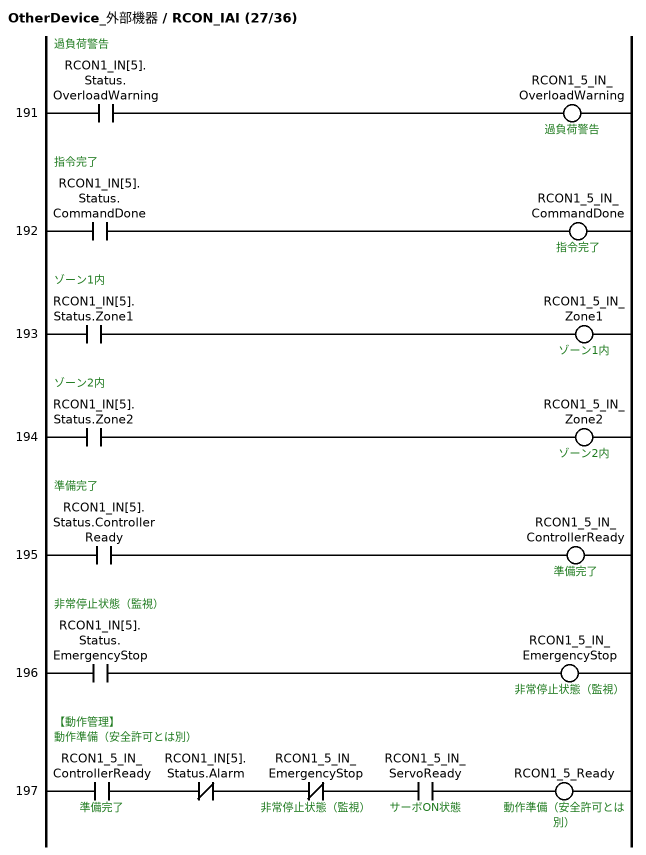
(* [picture p72: OtherDevice_外部機器 / RCON_IAI, rungs 191-197] *)
(* Rung 191: 過負荷警告 *)
RCON1_5_IN_OverloadWarning := RCON1_IN[5].Status.OverloadWarning;
(* Rung 192: 指令完了 *)
RCON1_5_IN_CommandDone := RCON1_IN[5].Status.CommandDone;
(* Rung 193: ゾーン1内 *)
RCON1_5_IN_Zone1 := RCON1_IN[5].Status.Zone1;
(* Rung 194: ゾーン2内 *)
RCON1_5_IN_Zone2 := RCON1_IN[5].Status.Zone2;
(* Rung 195: 準備完了 *)
RCON1_5_IN_ControllerReady := RCON1_IN[5].Status.ControllerReady;
(* Rung 196: 非常停止状態（監視） *)
RCON1_5_IN_EmergencyStop := RCON1_IN[5].Status.EmergencyStop;
(* Rung 197: 【動作管理】 / 動作準備（安全許可とは別） *)
RCON1_5_Ready := RCON1_5_IN_ControllerReady AND NOT RCON1_IN[5].Status.Alarm AND NOT RCON1_5_IN_EmergencyStop AND RCON1_5_IN_ServoReady;

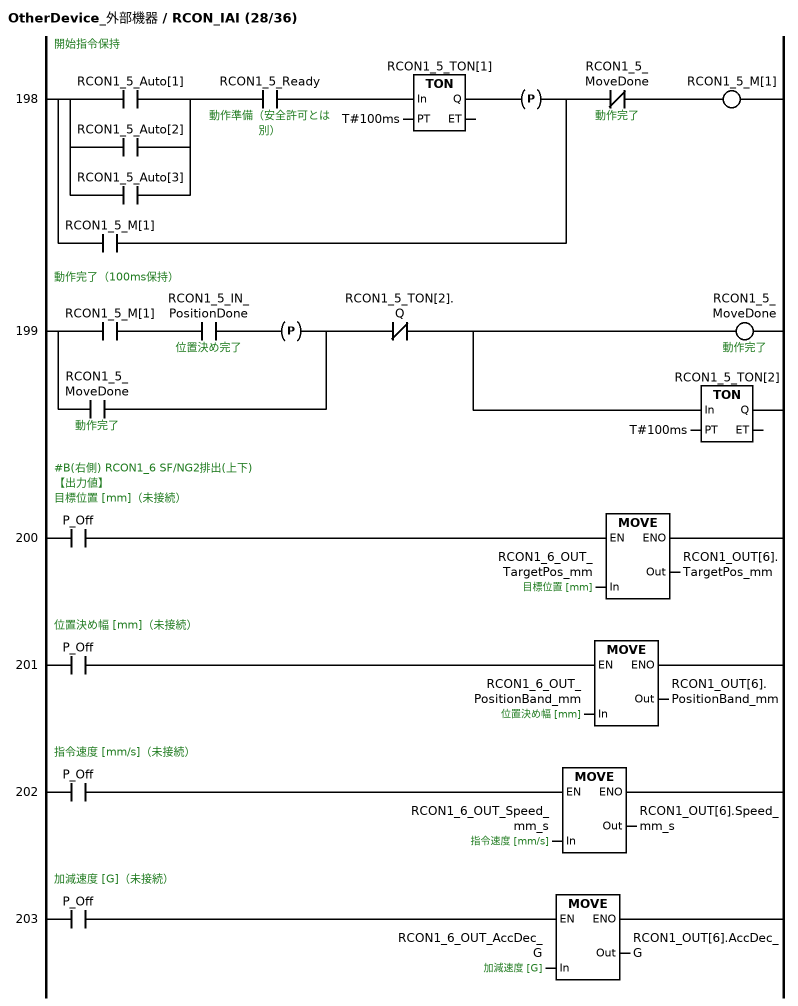
(* Rung 198: 開始指令保持 *)
RCON1_5_TON[1](In := (RCON1_5_Auto[1] OR RCON1_5_Auto[2] OR RCON1_5_Auto[3]) AND RCON1_5_Ready, PT := T#100ms);
_e18(CLK := RCON1_5_TON[1].Q);
RCON1_5_M[1] := (_e18.Q OR RCON1_5_M[1]) AND NOT RCON1_5_MoveDone;
(* Rung 199: 動作完了（100ms保持） *)
_e19(CLK := RCON1_5_M[1] AND RCON1_5_IN_PositionDone);
_p20 := (_e19.Q OR RCON1_5_MoveDone) AND NOT RCON1_5_TON[2].Q;
RCON1_5_MoveDone := _p20;
RCON1_5_TON[2](In := _p20, PT := T#100ms);
(* Rung 200: #B(右側) RCON1_6 SF/NG2排出(上下) / 【出力値】 / 目標位置 [mm]（未接続） *)
IF P_Off THEN RCON1_OUT[6].TargetPos_mm := RCON1_6_OUT_TargetPos_mm; END_IF;
(* Rung 201: 位置決め幅 [mm]（未接続） *)
IF P_Off THEN RCON1_OUT[6].PositionBand_mm := RCON1_6_OUT_PositionBand_mm; END_IF;
(* Rung 202: 指令速度 [mm/s]（未接続） *)
IF P_Off THEN RCON1_OUT[6].Speed_mm_s := RCON1_6_OUT_Speed_mm_s; END_IF;
(* Rung 203: 加減速度 [G]（未接続） *)
IF P_Off THEN RCON1_OUT[6].AccDec_G := RCON1_6_OUT_AccDec_G; END_IF;

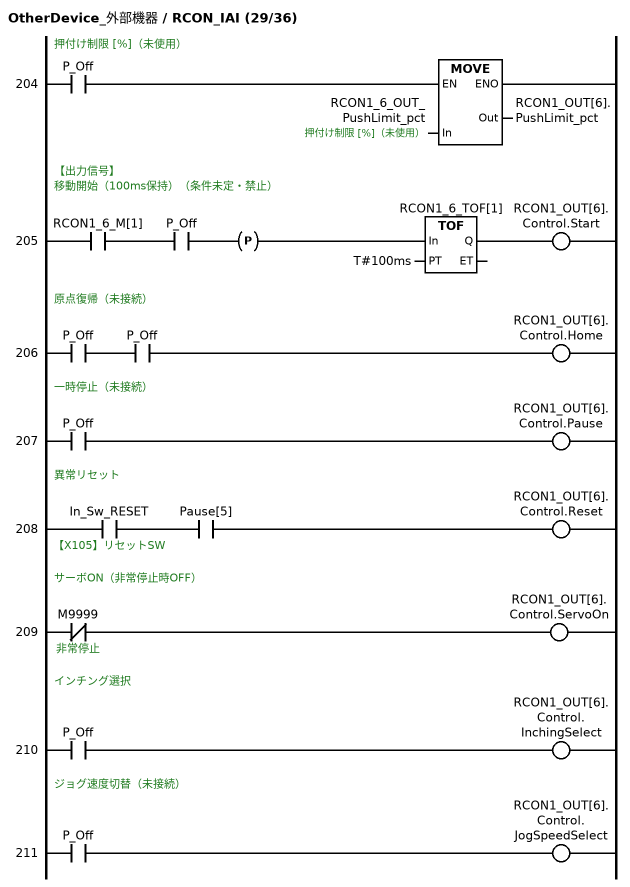
(* Rung 204: 押付け制限 [%]（未使用） *)
IF P_Off THEN RCON1_OUT[6].PushLimit_pct := RCON1_6_OUT_PushLimit_pct; END_IF;
(* Rung 205: 【出力信号】 / 移動開始（100ms保持）（条件未定・禁止） *)
_e21(CLK := RCON1_6_M[1] AND P_Off);
RCON1_6_TOF[1](In := _e21.Q, PT := T#100ms);
RCON1_OUT[6].Control.Start := RCON1_6_TOF[1].Q;
(* Rung 206: 原点復帰（未接続） *)
RCON1_OUT[6].Control.Home := P_Off AND P_Off;
(* Rung 207: 一時停止（未接続） *)
RCON1_OUT[6].Control.Pause := P_Off;
(* Rung 208: 異常リセット *)
RCON1_OUT[6].Control.Reset := In_Sw_RESET AND Pause[5];
(* Rung 209: サーボON（非常停止時OFF） *)
RCON1_OUT[6].Control.ServoOn := NOT M9999;
(* Rung 210: インチング選択 *)
RCON1_OUT[6].Control.InchingSelect := P_Off;
(* Rung 211: ジョグ速度切替（未接続） *)
RCON1_OUT[6].Control.JogSpeedSelect := P_Off;

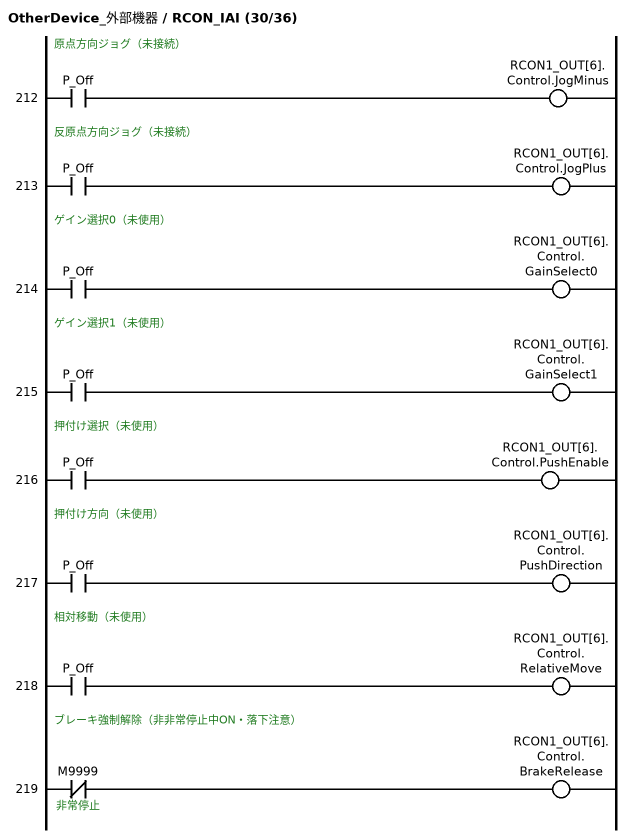
(* Rung 212: 原点方向ジョグ（未接続） *)
RCON1_OUT[6].Control.JogMinus := P_Off;
(* Rung 213: 反原点方向ジョグ（未接続） *)
RCON1_OUT[6].Control.JogPlus := P_Off;
(* Rung 214: ゲイン選択0（未使用） *)
RCON1_OUT[6].Control.GainSelect0 := P_Off;
(* Rung 215: ゲイン選択1（未使用） *)
RCON1_OUT[6].Control.GainSelect1 := P_Off;
(* Rung 216: 押付け選択（未使用） *)
RCON1_OUT[6].Control.PushEnable := P_Off;
(* Rung 217: 押付け方向（未使用） *)
RCON1_OUT[6].Control.PushDirection := P_Off;
(* Rung 218: 相対移動（未使用） *)
RCON1_OUT[6].Control.RelativeMove := P_Off;
(* Rung 219: ブレーキ強制解除（非非常停止中ON・落下注意） *)
RCON1_OUT[6].Control.BrakeRelease := NOT M9999;

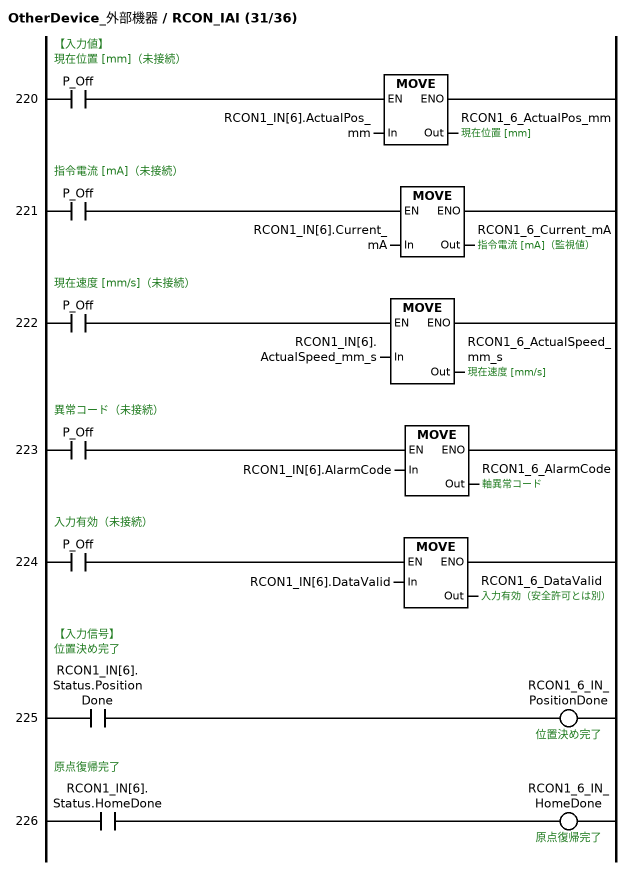
(* Rung 220: 【入力値】 / 現在位置 [mm]（未接続） *)
IF P_Off THEN RCON1_6_ActualPos_mm := RCON1_IN[6].ActualPos_mm; END_IF;
(* Rung 221: 指令電流 [mA]（未接続） *)
IF P_Off THEN RCON1_6_Current_mA := RCON1_IN[6].Current_mA; END_IF;
(* Rung 222: 現在速度 [mm/s]（未接続） *)
IF P_Off THEN RCON1_6_ActualSpeed_mm_s := RCON1_IN[6].ActualSpeed_mm_s; END_IF;
(* Rung 223: 異常コード（未接続） *)
IF P_Off THEN RCON1_6_AlarmCode := RCON1_IN[6].AlarmCode; END_IF;
(* Rung 224: 入力有効（未接続） *)
IF P_Off THEN RCON1_6_DataValid := RCON1_IN[6].DataValid; END_IF;
(* Rung 225: 【入力信号】 / 位置決め完了 *)
RCON1_6_IN_PositionDone := RCON1_IN[6].Status.PositionDone;
(* Rung 226: 原点復帰完了 *)
RCON1_6_IN_HomeDone := RCON1_IN[6].Status.HomeDone;

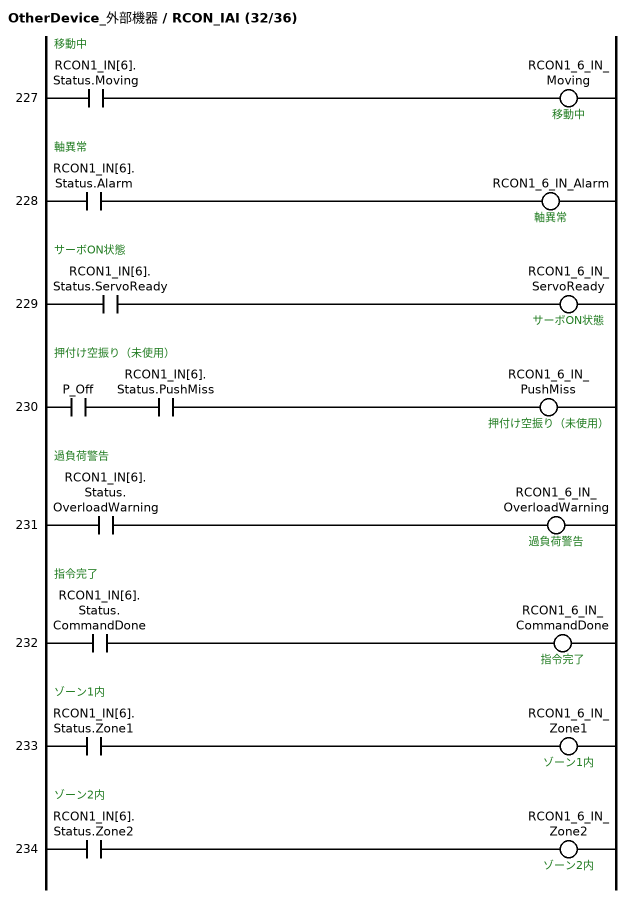
(* Rung 227: 移動中 *)
RCON1_6_IN_Moving := RCON1_IN[6].Status.Moving;
(* Rung 228: 軸異常 *)
RCON1_6_IN_Alarm := RCON1_IN[6].Status.Alarm;
(* Rung 229: サーボON状態 *)
RCON1_6_IN_ServoReady := RCON1_IN[6].Status.ServoReady;
(* Rung 230: 押付け空振り（未使用） *)
RCON1_6_IN_PushMiss := P_Off AND RCON1_IN[6].Status.PushMiss;
(* Rung 231: 過負荷警告 *)
RCON1_6_IN_OverloadWarning := RCON1_IN[6].Status.OverloadWarning;
(* Rung 232: 指令完了 *)
RCON1_6_IN_CommandDone := RCON1_IN[6].Status.CommandDone;
(* Rung 233: ゾーン1内 *)
RCON1_6_IN_Zone1 := RCON1_IN[6].Status.Zone1;
(* Rung 234: ゾーン2内 *)
RCON1_6_IN_Zone2 := RCON1_IN[6].Status.Zone2;

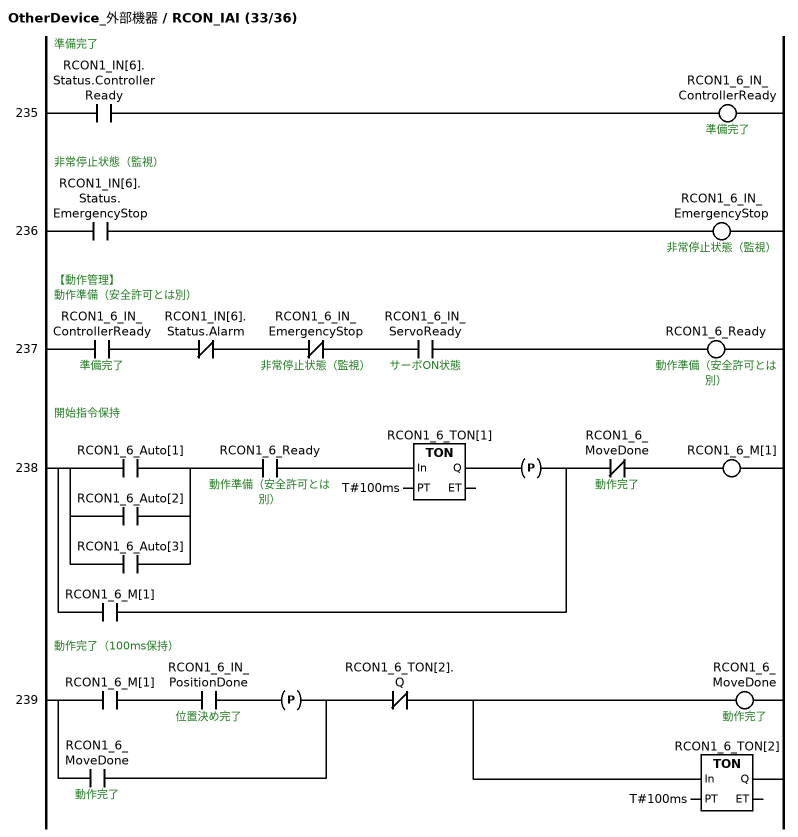
(* Rung 235: 準備完了 *)
RCON1_6_IN_ControllerReady := RCON1_IN[6].Status.ControllerReady;
(* Rung 236: 非常停止状態（監視） *)
RCON1_6_IN_EmergencyStop := RCON1_IN[6].Status.EmergencyStop;
(* Rung 237: 【動作管理】 / 動作準備（安全許可とは別） *)
RCON1_6_Ready := RCON1_6_IN_ControllerReady AND NOT RCON1_IN[6].Status.Alarm AND NOT RCON1_6_IN_EmergencyStop AND RCON1_6_IN_ServoReady;
(* Rung 238: 開始指令保持 *)
RCON1_6_TON[1](In := (RCON1_6_Auto[1] OR RCON1_6_Auto[2] OR RCON1_6_Auto[3]) AND RCON1_6_Ready, PT := T#100ms);
_e22(CLK := RCON1_6_TON[1].Q);
RCON1_6_M[1] := (_e22.Q OR RCON1_6_M[1]) AND NOT RCON1_6_MoveDone;
(* Rung 239: 動作完了（100ms保持） *)
_e23(CLK := RCON1_6_M[1] AND RCON1_6_IN_PositionDone);
_p24 := (_e23.Q OR RCON1_6_MoveDone) AND NOT RCON1_6_TON[2].Q;
RCON1_6_MoveDone := _p24;
RCON1_6_TON[2](In := _p24, PT := T#100ms);

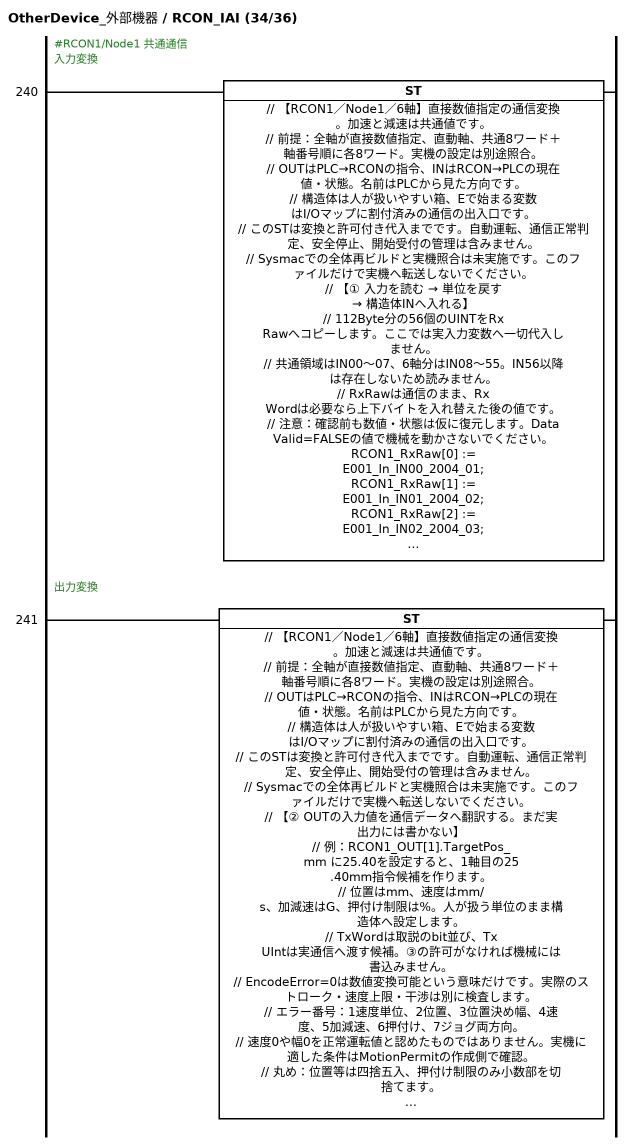
(* Rung 240: #RCON1/Node1 共通通信 / 入力変換 *)
// 【RCON1／Node1／6軸】直接数値指定の通信変換。加速と減速は共通値です。
// 前提：全軸が直接数値指定、直動軸、共通8ワード＋軸番号順に各8ワード。実機の設定は別途照合。
// OUTはPLC→RCONの指令、INはRCON→PLCの現在値・状態。名前はPLCから見た方向です。
// 構造体は人が扱いやすい箱、Eで始まる変数はI/Oマップに割付済みの通信の出入口です。
// このSTは変換と許可付き代入までです。自動運転、通信正常判定、安全停止、開始受付の管理は含みません。
// Sysmacでの全体再ビルドと実機照合は未実施です。このファイルだけで実機へ転送しないでください。
// 【① 入力を読む → 単位を戻す → 構造体INへ入れる】
// 112Byte分の56個のUINTをRxRawへコピーします。ここでは実入力変数へ一切代入しません。
// 共通領域はIN00～07、6軸分はIN08～55。IN56以降は存在しないため読みません。
// RxRawは通信のまま、RxWordは必要なら上下バイトを入れ替えた後の値です。
// 注意：確認前も数値・状態は仮に復元します。DataValid=FALSEの値で機械を動かさないでください。
RCON1_RxRaw[0] := E001_In_IN00_2004_01;
RCON1_RxRaw[1] := E001_In_IN01_2004_02;
RCON1_RxRaw[2] := E001_In_IN02_2004_03;
RCON1_RxRaw[3] := E001_In_IN03_2004_04;
RCON1_RxRaw[4] := E001_In_IN04_2004_05;
RCON1_RxRaw[5] := E001_In_IN05_2004_06;
RCON1_RxRaw[6] := E001_In_IN06_2004_07;
RCON1_RxRaw[7] := E001_In_IN07_2004_08;
RCON1_RxRaw[8] := E001_In_IN08_2004_09;
RCON1_RxRaw[9] := E001_In_IN09_2004_0A;
RCON1_RxRaw[10] := E001_In_IN10_2004_0B;
RCON1_RxRaw[11] := E001_In_IN11_2004_0C;
RCON1_RxRaw[12] := E001_In_IN12_2004_0D;
RCON1_RxRaw[13] := E001_In_IN13_2004_0E;
RCON1_RxRaw[14] := E001_In_IN14_2004_0F;
RCON1_RxRaw[15] := E001_In_IN15_2004_10;
RCON1_RxRaw[16] := E001_In_IN16_2004_11;
RCON1_RxRaw[17] := E001_In_IN17_2004_12;
RCON1_RxRaw[18] := E001_In_IN18_2004_13;
RCON1_RxRaw[19] := E001_In_IN19_2004_14;
RCON1_RxRaw[20] := E001_In_IN20_2004_15;
RCON1_RxRaw[21] := E001_In_IN21_2004_16;
RCON1_RxRaw[22] := E001_In_IN22_2004_17;
RCON1_RxRaw[23] := E001_In_IN23_2004_18;
RCON1_RxRaw[24] := E001_In_IN24_2004_19;
RCON1_RxRaw[25] := E001_In_IN25_2004_1A;
RCON1_RxRaw[26] := E001_In_IN26_2004_1B;
RCON1_RxRaw[27] := E001_In_IN27_2004_1C;
RCON1_RxRaw[28] := E001_In_IN28_2004_1D;
RCON1_RxRaw[29] := E001_In_IN29_2004_1E;
RCON1_RxRaw[30] := E001_In_IN30_2004_1F;
RCON1_RxRaw[31] := E001_In_IN31_2004_20;
RCON1_RxRaw[32] := E001_In_IN32_2004_21;
RCON1_RxRaw[33] := E001_In_IN33_2004_22;
RCON1_RxRaw[34] := E001_In_IN34_2004_23;
RCON1_RxRaw[35] := E001_In_IN35_2004_24;
RCON1_RxRaw[36] := E001_In_IN36_2004_25;
RCON1_RxRaw[37] := E001_In_IN37_2004_26;
RCON1_RxRaw[38] := E001_In_IN38_2004_27;
RCON1_RxRaw[39] := E001_In_IN39_2004_28;
RCON1_RxRaw[40] := E001_In_IN40_2004_29;
RCON1_RxRaw[41] := E001_In_IN41_2004_2A;
RCON1_RxRaw[42] := E001_In_IN42_2004_2B;
RCON1_RxRaw[43] := E001_In_IN43_2004_2C;
RCON1_RxRaw[44] := E001_In_IN44_2004_2D;
RCON1_RxRaw[45] := E001_In_IN45_2004_2E;
RCON1_RxRaw[46] := E001_In_IN46_2004_2F;
RCON1_RxRaw[47] := E001_In_IN47_2004_30;
RCON1_RxRaw[48] := E001_In_IN48_2004_31;
RCON1_RxRaw[49] := E001_In_IN49_2004_32;
RCON1_RxRaw[50] := E001_In_IN50_2004_33;
RCON1_RxRaw[51] := E001_In_IN51_2004_34;
RCON1_RxRaw[52] := E001_In_IN52_2004_35;
RCON1_RxRaw[53] := E001_In_IN53_2004_36;
RCON1_RxRaw[54] := E001_In_IN54_2004_37;
RCON1_RxRaw[55] := E001_In_IN55_2004_38;
// 取説の論理ワードへ正規化。Swapは1ワード内の上下バイト交換です。
// SwapBytesは推測で設定せず、既知の位置とbitで実機照合してください。
FOR ConvWordIndex := INT#0 TO INT#55 DO
    RCON1_RxWord[ConvWordIndex] := UINT_TO_WORD(RCON1_RxRaw[ConvWordIndex]);
    IF RCON1_SwapBytes THEN
        RCON1_RxWord[ConvWordIndex] := Swap(RCON1_RxWord[ConvWordIndex]);
    END_IF;
END_FOR;

ConvUnitOK := (RCON1_SpeedUnit_mm_s = LREAL#1.0) OR
              (RCON1_SpeedUnit_mm_s = LREAL#0.1);

// 【①-2 共通状態】IN00はユニット全体、IN01は各軸のリンク情報です。
// TestABit(ワード, bit番号)は、そのスイッチがONかをBOOLで取り出す命令です。
// 例：IN01のb0は軸No.0→配列[1]、b1は軸No.1→配列[2]。配列番号と実機軸番号は1違います。
// 共通固定領域。ここで使うbit番号は取説の論理bitです（MJ0384 6-24～6-25）。
RCON1_GwRun := TestABit(RCON1_RxWord[0], USINT#15);
RCON1_GwControllerCommLatch := TestABit(RCON1_RxWord[0], USINT#14);
RCON1_GwAxisCommError := TestABit(RCON1_RxWord[0], USINT#13);
RCON1_GwManual := TestABit(RCON1_RxWord[0], USINT#12);
RCON1_GwHeavyAlarm := TestABit(RCON1_RxWord[0], USINT#11);
RCON1_GwLightAlarm := TestABit(RCON1_RxWord[0], USINT#10);
RCON1_GwSystemStop := TestABit(RCON1_RxWord[0], USINT#8);
RCON1_GwAlarmCode := WORD_TO_UINT(RCON1_RxWord[0] AND WORD#16#00FF);
FOR ConvWordIndex := INT#0 TO INT#4 DO
    RCON1_PowerStateRaw[ConvWordIndex] := RCON1_RxWord[ConvWordIndex + INT#2];
END_FOR;

// 【①-3 軸ごとに同じ読取りを繰り返す】
// FORは1～6軸を順番に処理します。ConvBaseはその軸の先頭番号です。
// 計算：8+(軸番号-1)×8。1軸目=8、2軸目=16、3軸目=24。先頭8ワードは共通領域です。
FOR ConvAxisIndex := INT#1 TO INT#6 DO
    ConvBase := INT#8 + (ConvAxisIndex - INT#1) * INT#8;
    RCON1_AxisLinked[ConvAxisIndex] :=
        TestABit(RCON1_RxWord[1], INT_TO_USINT(ConvAxisIndex - INT#1));

// 例：下位2540／上位0なら32bit値2540→25.40mm。
// 上位を16bit左に動かして下位とORで重ねます。SHLが左シフト、ORがビットの合成です。
// 負位置はDWORD_TO_DINTで符号を復元。下位62996／上位65535なら-2540→-25.40mm。
    // 現在位置：下位・上位を結合、符号付き32bitとして解釈、0.01mmをmmへ。
    ConvDWord := SHL(WORD_TO_DWORD(RCON1_RxWord[ConvBase + INT#1]), ULINT#16)
                 OR WORD_TO_DWORD(RCON1_RxWord[ConvBase]);
    RCON1_IN[ConvAxisIndex].ActualPos_mm :=
        DINT_TO_LREAL(DWORD_TO_DINT(ConvDWord)) * LREAL#0.01;

    // 電流：32bitのmA。RCON-PCでは指令電流であり、実測トルクではありません。
    ConvDWord := SHL(WORD_TO_DWORD(RCON1_RxWord[ConvBase + INT#3]), ULINT#16)
                 OR WORD_TO_DWORD(RCON1_RxWord[ConvBase + INT#2]);
    RCON1_IN[ConvAxisIndex].Current_mA := DWORD_TO_DINT(ConvDWord);

    // 現在速度：16bitの負数をINTとして読む。UINTのまま速度にしません。
    IF ConvUnitOK THEN
        RCON1_IN[ConvAxisIndex].ActualSpeed_mm_s :=
            INT_TO_LREAL(WORD_TO_INT(RCON1_RxWord[ConvBase + INT#4])) * RCON1_SpeedUnit_mm_s;
    END_IF;
    // 単位不明のとき速度は前値を保持し、DataValidはFALSEにします。
    // 軸内の+5ワードは予約のため値を使用しません。
    RCON1_IN[ConvAxisIndex].AlarmCode := WORD_TO_UINT(RCON1_RxWord[ConvBase + INT#6]);

// 例：Status.ServoReady=TRUEは「サーボON状態を受信した」という意味。
// OUT側Control.ServoOn=TRUEは「サーボONを要求する」という意味で、指令と結果を区別します。
    // 状態ワード：12個のBOOLへ分解。予約b6,b9～11は使いません。
    RCON1_IN[ConvAxisIndex].Status.PositionDone := TestABit(RCON1_RxWord[ConvBase + INT#7], USINT#0);
    RCON1_IN[ConvAxisIndex].Status.HomeDone := TestABit(RCON1_RxWord[ConvBase + INT#7], USINT#1);
    RCON1_IN[ConvAxisIndex].Status.Moving := TestABit(RCON1_RxWord[ConvBase + INT#7], USINT#2);
    RCON1_IN[ConvAxisIndex].Status.Alarm := TestABit(RCON1_RxWord[ConvBase + INT#7], USINT#3);
    RCON1_IN[ConvAxisIndex].Status.ServoReady := TestABit(RCON1_RxWord[ConvBase + INT#7], USINT#4);
    RCON1_IN[ConvAxisIndex].Status.PushMiss := TestABit(RCON1_RxWord[ConvBase + INT#7], USINT#5);
    RCON1_IN[ConvAxisIndex].Status.OverloadWarning := TestABit(RCON1_RxWord[ConvBase + INT#7], USINT#7);
    RCON1_IN[ConvAxisIndex].Status.CommandDone := TestABit(RCON1_RxWord[ConvBase + INT#7], USINT#8);
    RCON1_IN[ConvAxisIndex].Status.Zone1 := TestABit(RCON1_RxWord[ConvBase + INT#7], USINT#12);
    RCON1_IN[ConvAxisIndex].Status.Zone2 := TestABit(RCON1_RxWord[ConvBase + INT#7], USINT#13);
    RCON1_IN[ConvAxisIndex].Status.ControllerReady := TestABit(RCON1_RxWord[ConvBase + INT#7], USINT#14);
    RCON1_IN[ConvAxisIndex].Status.EmergencyStop := TestABit(RCON1_RxWord[ConvBase + INT#7], USINT#15);

    // DataValidは直接受信bitではなく、今回の内部設計で決めた内部判定です。
    // CommOKはCPUの実通信状態から別途作成。単にTRUE固定にしないでください。
    // DataValidは運転許可や安全保証ではありません。各異常・原点等は別途確認。
    RCON1_IN[ConvAxisIndex].DataValid := RCON1_CommOK AND RCON1_LayoutConfirmed
        AND RCON1_ByteOrderConfirmed AND ConvUnitOK AND RCON1_GwRun
        AND RCON1_AxisLinked[ConvAxisIndex] AND NOT RCON1_GwAxisCommError;
END_FOR;
(* Rung 241: 出力変換 *)
// 【RCON1／Node1／6軸】直接数値指定の通信変換。加速と減速は共通値です。
// 前提：全軸が直接数値指定、直動軸、共通8ワード＋軸番号順に各8ワード。実機の設定は別途照合。
// OUTはPLC→RCONの指令、INはRCON→PLCの現在値・状態。名前はPLCから見た方向です。
// 構造体は人が扱いやすい箱、Eで始まる変数はI/Oマップに割付済みの通信の出入口です。
// このSTは変換と許可付き代入までです。自動運転、通信正常判定、安全停止、開始受付の管理は含みません。
// Sysmacでの全体再ビルドと実機照合は未実施です。このファイルだけで実機へ転送しないでください。
// 【② OUTの入力値を通信データへ翻訳する。まだ実出力には書かない】
// 例：RCON1_OUT[1].TargetPos_mm に25.40を設定すると、1軸目の25.40mm指令候補を作ります。
// 位置はmm、速度はmm/s、加減速はG、押付け制限は%。人が扱う単位のまま構造体へ設定します。
// TxWordは取説のbit並び、TxUIntは実通信へ渡す候補。③の許可がなければ機械には書込みません。
// EncodeError=0は数値変換可能という意味だけです。実際のストローク・速度上限・干渉は別に検査します。
// エラー番号：1速度単位、2位置、3位置決め幅、4速度、5加減速、6押付け、7ジョグ両方向。
// 速度0や幅0を正常運転値と認めたものではありません。実機に適した条件はMotionPermitの作成側で確認。
// 丸め：位置等は四捨五入、押付け制限のみ小数部を切捨てます。

ConvUnitOK := (RCON1_SpeedUnit_mm_s = LREAL#1.0) OR
              (RCON1_SpeedUnit_mm_s = LREAL#0.1);

// 共通制御：MONは論理b15、RTEは論理b13。他のbitは0。
// MONを落とす処理を安全停止として扱わないでください。
RCON1_TxWord[0] := WORD#16#0000;
IF RCON1_GwMON_Request THEN
    RCON1_TxWord[0] := RCON1_TxWord[0] OR WORD#16#8000;
END_IF;
IF RCON1_GwRTE_Request THEN
    RCON1_TxWord[0] := RCON1_TxWord[0] OR WORD#16#2000;
END_IF;

FOR ConvAxisIndex := INT#1 TO INT#6 DO
    ConvBase := INT#8 + (ConvAxisIndex - INT#1) * INT#8;
    RCON1_EncodeError[ConvAxisIndex] := UINT#0;

    // 比較で範囲を確認してから型変換するため、NaN・無限大も変換対象から外れます。
    // 位置・幅9999.99mmはこの案で採用する通信範囲の上限で、実機ストロークではありません。
    IF NOT ConvUnitOK THEN
        RCON1_EncodeError[ConvAxisIndex] := UINT#1;
    ELSIF NOT ((RCON1_OUT[ConvAxisIndex].TargetPos_mm >= LREAL#-9999.99) AND
               (RCON1_OUT[ConvAxisIndex].TargetPos_mm <= LREAL#9999.99)) THEN
        RCON1_EncodeError[ConvAxisIndex] := UINT#2;
    ELSIF NOT ((RCON1_OUT[ConvAxisIndex].PositionBand_mm >= LREAL#0.0) AND
               (RCON1_OUT[ConvAxisIndex].PositionBand_mm <= LREAL#9999.99)) THEN
        RCON1_EncodeError[ConvAxisIndex] := UINT#3;
    ELSIF NOT ((RCON1_OUT[ConvAxisIndex].Speed_mm_s >= LREAL#0.0) AND
               (RCON1_OUT[ConvAxisIndex].Speed_mm_s <= LREAL#65535.0 * RCON1_SpeedUnit_mm_s)) THEN
        RCON1_EncodeError[ConvAxisIndex] := UINT#4;
    ELSIF NOT ((RCON1_OUT[ConvAxisIndex].AccDec_G >= LREAL#0.0) AND
               (RCON1_OUT[ConvAxisIndex].AccDec_G <= LREAL#655.35)) THEN
        RCON1_EncodeError[ConvAxisIndex] := UINT#5;
    ELSIF NOT ((RCON1_OUT[ConvAxisIndex].PushLimit_pct >= LREAL#0.0) AND
               (RCON1_OUT[ConvAxisIndex].PushLimit_pct <= LREAL#200.0)) THEN
        RCON1_EncodeError[ConvAxisIndex] := UINT#6;
    ELSIF RCON1_OUT[ConvAxisIndex].Control.JogMinus AND RCON1_OUT[ConvAxisIndex].Control.JogPlus THEN
        RCON1_EncodeError[ConvAxisIndex] := UINT#7;
    END_IF;

    RCON1_EncodeOK[ConvAxisIndex] := RCON1_EncodeError[ConvAxisIndex] = UINT#0;
    IF RCON1_EncodeOK[ConvAxisIndex] THEN
    // 【数値例】TargetPos_mm=25.40→×100で2540。下位ワード2540、上位ワード0。
// 700.25mm→70025なので下位4489、上位1。65536を超えた分が上位に入ります。
// DINTは符号付きの数、DWORDは同じ32bitの模様。負数の符号を壊さず分割するために使い分けます。
// TRUNCは小数部を捨てます。正数+0.5／負数-0.5を先に行い、四捨五入を明示しています。
    // 目標位置：mmから0.01mmの符号付き整数へ。
        ConvScaled := RCON1_OUT[ConvAxisIndex].TargetPos_mm * LREAL#100.0;
        IF ConvScaled >= LREAL#0.0 THEN
            ConvPos := LINT_TO_DINT(TRUNC(ConvScaled + LREAL#0.5));
        ELSE
            ConvPos := LINT_TO_DINT(TRUNC(ConvScaled - LREAL#0.5));
        END_IF;
        // 負数を含む32bitパターンを保ち、下位・上位の16bitへ分割。
        ConvDWord := DINT_TO_DWORD(ConvPos);
        RCON1_TxWord[ConvBase] := DWORD_TO_WORD(ConvDWord AND DWORD#16#0000FFFF);
        RCON1_TxWord[ConvBase + INT#1] := DWORD_TO_WORD(SHR(ConvDWord, ULINT#16));

        // 位置決め幅：非負の内部整数としてUDINTを選定（メーカーの符号なし保証ではありません）。
        ConvBand := LINT_TO_UDINT(TRUNC(RCON1_OUT[ConvAxisIndex].PositionBand_mm * LREAL#100.0 + LREAL#0.5));
        ConvDWord := UDINT_TO_DWORD(ConvBand);
        RCON1_TxWord[ConvBase + INT#2] := DWORD_TO_WORD(ConvDWord AND DWORD#16#0000FFFF);
        RCON1_TxWord[ConvBase + INT#3] := DWORD_TO_WORD(SHR(ConvDWord, ULINT#16));

// 速度20mm/s：速度単位1.0なら20、0.1なら200を送信します。
// 加減速0.20G：×100して20。加速と減速の両方に同じ値を使います。
// 押付け50%：×255÷100=127.5を切捨てて127。押付けの使用可否・上限は実機仕様で別確認。
        // 速度は1カウント量が1.0か0.1かで値が10倍変わります。
        ConvSpeed := LINT_TO_UINT(TRUNC(RCON1_OUT[ConvAxisIndex].Speed_mm_s / RCON1_SpeedUnit_mm_s + LREAL#0.5));
        ConvAccDec := LINT_TO_UINT(TRUNC(RCON1_OUT[ConvAxisIndex].AccDec_G * LREAL#100.0 + LREAL#0.5));
        ConvPush := LINT_TO_UINT(TRUNC(RCON1_OUT[ConvAxisIndex].PushLimit_pct * LREAL#255.0 / LREAL#100.0));
        RCON1_TxWord[ConvBase + INT#4] := UINT_TO_WORD(ConvSpeed);
        RCON1_TxWord[ConvBase + INT#5] := UINT_TO_WORD(ConvAccDec);
        RCON1_TxWord[ConvBase + INT#6] := UINT_TO_WORD(ConvPush);
    END_IF;
    // 不正値の場合、数値ワードは前値保持。EncodeOK=FALSEで03の書込みを抑止。
    // 前値保持は停止指令ではありません。停止・異常処理は別途設計してください。

    // Controlを論理bitへ詰める。予約b9は必ず0。
    RCON1_TxWord[ConvBase + INT#7] := WORD#16#0000;
// b0 DSTR／Control.Start：TRUEで開始要求。受付応答と10ms以上の保持を確認してOFF。常時ONにしない。
    IF RCON1_OUT[ConvAxisIndex].Control.Start THEN
        RCON1_TxWord[ConvBase + INT#7] := RCON1_TxWord[ConvBase + INT#7] OR WORD#16#0001;
    END_IF;
// b1 HOME／Control.Home：TRUEで原点復帰を指令。原点復帰完了はIN側HomeDoneで確認。
    IF RCON1_OUT[ConvAxisIndex].Control.Home THEN
        RCON1_TxWord[ConvBase + INT#7] := RCON1_TxWord[ConvBase + INT#7] OR WORD#16#0002;
    END_IF;
// b2 STP／Control.Pause：TRUEで一時停止、FALSEで解除。非常停止・安全停止の代用ではない。
    IF RCON1_OUT[ConvAxisIndex].Control.Pause THEN
        RCON1_TxWord[ConvBase + INT#7] := RCON1_TxWord[ConvBase + INT#7] OR WORD#16#0004;
    END_IF;
// b3 RES／Control.Reset：TRUEでアラームリセット要求。コールドスタート級の異常には使用できない。
    IF RCON1_OUT[ConvAxisIndex].Control.Reset THEN
        RCON1_TxWord[ConvBase + INT#7] := RCON1_TxWord[ConvBase + INT#7] OR WORD#16#0008;
    END_IF;
// b4 SON／Control.ServoOn：TRUEでサーボON要求。ON状態はIN側ServoReadyで確認。
    IF RCON1_OUT[ConvAxisIndex].Control.ServoOn THEN
        RCON1_TxWord[ConvBase + INT#7] := RCON1_TxWord[ConvBase + INT#7] OR WORD#16#0010;
    END_IF;
// b5 JISL／Control.InchingSelect：TRUEは一定距離のインチング、FALSEは押している間のジョグ。
    IF RCON1_OUT[ConvAxisIndex].Control.InchingSelect THEN
        RCON1_TxWord[ConvBase + INT#7] := RCON1_TxWord[ConvBase + INT#7] OR WORD#16#0020;
    END_IF;
// b6 JVEL／Control.JogSpeedSelect：FALSEは速度No.26・距離No.48、TRUEは速度No.47または指令速度・距離No.49。
    IF RCON1_OUT[ConvAxisIndex].Control.JogSpeedSelect THEN
        RCON1_TxWord[ConvBase + INT#7] := RCON1_TxWord[ConvBase + INT#7] OR WORD#16#0040;
    END_IF;
// b7 JOG-／Control.JogMinus：TRUEで原点方向へジョグ。反対方向指令との同時ONを防ぐ。
    IF RCON1_OUT[ConvAxisIndex].Control.JogMinus THEN
        RCON1_TxWord[ConvBase + INT#7] := RCON1_TxWord[ConvBase + INT#7] OR WORD#16#0080;
    END_IF;
// b8 JOG+／Control.JogPlus：TRUEで反原点方向へジョグ。反対方向指令との同時ONを防ぐ。
    IF RCON1_OUT[ConvAxisIndex].Control.JogPlus THEN
        RCON1_TxWord[ConvBase + INT#7] := RCON1_TxWord[ConvBase + INT#7] OR WORD#16#0100;
    END_IF;
// b10 GSL0／Control.GainSelect0：GainSelect1と組合せてサーボゲインセット0～3を選ぶ。機械調整用。
    IF RCON1_OUT[ConvAxisIndex].Control.GainSelect0 THEN
        RCON1_TxWord[ConvBase + INT#7] := RCON1_TxWord[ConvBase + INT#7] OR WORD#16#0400;
    END_IF;
// b11 GSL1／Control.GainSelect1：GainSelect0との2bitで選択。速度指令とは別の機能。
    IF RCON1_OUT[ConvAxisIndex].Control.GainSelect1 THEN
        RCON1_TxWord[ConvBase + INT#7] := RCON1_TxWord[ConvBase + INT#7] OR WORD#16#0800;
    END_IF;
// b12 PUSH／Control.PushEnable：TRUEは押付け、FALSEは通常位置決め。押付け条件は別途確認。
    IF RCON1_OUT[ConvAxisIndex].Control.PushEnable THEN
        RCON1_TxWord[ConvBase + INT#7] := RCON1_TxWord[ConvBase + INT#7] OR WORD#16#1000;
    END_IF;
// b13 DIR／Control.PushDirection：CON方式押付け時、TRUEは反原点方向、FALSEは原点方向。
    IF RCON1_OUT[ConvAxisIndex].Control.PushDirection THEN
        RCON1_TxWord[ConvBase + INT#7] := RCON1_TxWord[ConvBase + INT#7] OR WORD#16#2000;
    END_IF;
// b14 INC／Control.RelativeMove：FALSEは絶対座標、TRUEは現在位置からの相対移動量。
    IF RCON1_OUT[ConvAxisIndex].Control.RelativeMove THEN
        RCON1_TxWord[ConvBase + INT#7] := RCON1_TxWord[ConvBase + INT#7] OR WORD#16#4000;
    END_IF;
// b15 BKRL／Control.BrakeRelease：TRUEはブレーキ強制解除。通常FALSE。縦軸では落下等の危険がある。
    IF RCON1_OUT[ConvAxisIndex].Control.BrakeRelease THEN
        RCON1_TxWord[ConvBase + INT#7] := RCON1_TxWord[ConvBase + INT#7] OR WORD#16#8000;
    END_IF;
END_FOR;

// 論理ワードから実際に送るUINTへ。INと同じ1ワード内のバイト交換を適用します。
FOR ConvWordIndex := INT#0 TO INT#55 DO
    ConvWord := RCON1_TxWord[ConvWordIndex];
    IF RCON1_SwapBytes THEN
        ConvWord := Swap(ConvWord);
    END_IF;
    RCON1_TxUInt[ConvWordIndex] := WORD_TO_UINT(ConvWord);
END_FOR;

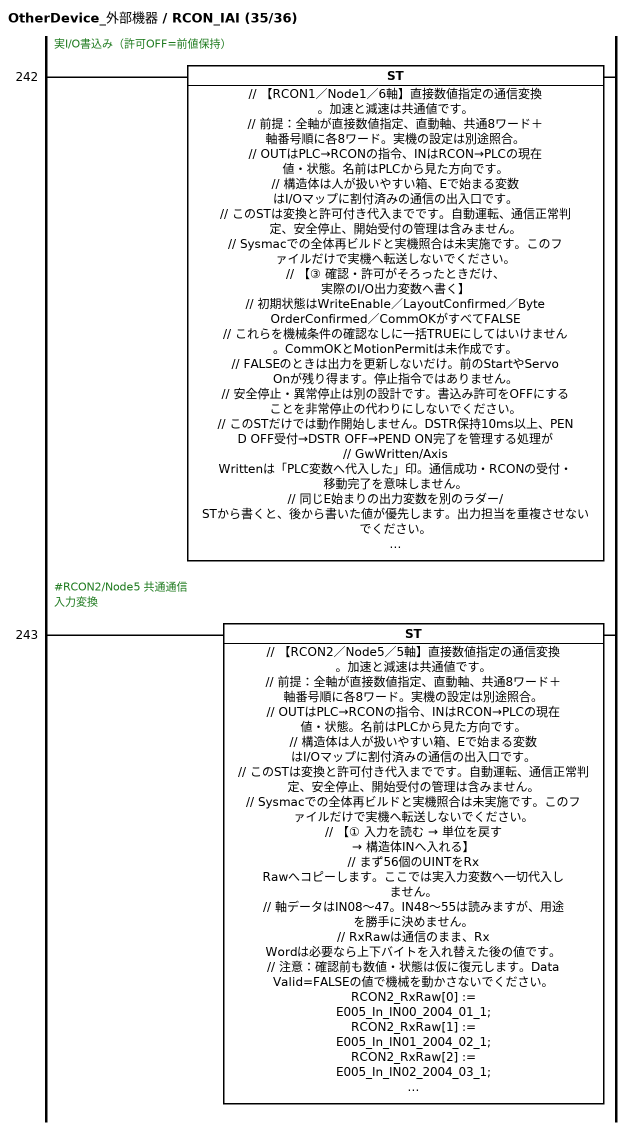
(* Rung 242: 実I/O書込み（許可OFF=前値保持） *)
// 【RCON1／Node1／6軸】直接数値指定の通信変換。加速と減速は共通値です。
// 前提：全軸が直接数値指定、直動軸、共通8ワード＋軸番号順に各8ワード。実機の設定は別途照合。
// OUTはPLC→RCONの指令、INはRCON→PLCの現在値・状態。名前はPLCから見た方向です。
// 構造体は人が扱いやすい箱、Eで始まる変数はI/Oマップに割付済みの通信の出入口です。
// このSTは変換と許可付き代入までです。自動運転、通信正常判定、安全停止、開始受付の管理は含みません。
// Sysmacでの全体再ビルドと実機照合は未実施です。このファイルだけで実機へ転送しないでください。
// 【③ 確認・許可がそろったときだけ、実際のI/O出力変数へ書く】
// 初期状態はWriteEnable／LayoutConfirmed／ByteOrderConfirmed／CommOKがすべてFALSEです。
// これらを機械条件の確認なしに一括TRUEにしてはいけません。CommOKとMotionPermitは未作成です。
// FALSEのときは出力を更新しないだけ。前のStartやServoOnが残り得ます。停止指令ではありません。
// 安全停止・異常停止は別の設計です。書込み許可をOFFにすることを非常停止の代わりにしないでください。
// このSTだけでは動作開始しません。DSTR保持10ms以上、PEND OFF受付→DSTR OFF→PEND ON完了を管理する処理が必要です。
// GwWritten/AxisWrittenは「PLC変数へ代入した」印。通信成功・RCONの受付・移動完了を意味しません。
// 同じE始まりの出力変数を別のラダー/STから書くと、後から書いた値が優先します。出力担当を重複させないでください。

RCON1_GwWritten := FALSE;
FOR ConvAxisIndex := INT#1 TO INT#6 DO
    RCON1_AxisWritten[ConvAxisIndex] := FALSE;
END_FOR;

IF RCON1_WriteEnable AND RCON1_LayoutConfirmed AND RCON1_ByteOrderConfirmed AND RCON1_CommOK THEN
// 共通指令はMON/RTEのみ。最初のRUN応答に必要なため、軸DataValidとは別にGwApplyで許可します。
    IF RCON1_GwApply THEN
        E001_Out_OUT00_2003_01 := RCON1_TxUInt[0];
        RCON1_GwWritten := TRUE;
    END_IF;

// 1軸目＝実機軸No.0。OUT08～OUT15の8ワードをまとめて代入。
// AxisApply=この軸の更新許可、EncodeOK=変換OK、DataValid=入力情報の条件確認、MotionPermit=機械側の運転許可。
// 途中1ワードだけではなく、位置・幅・速度・加減速・押付け・制御を一組として渡します。
    IF RCON1_AxisApply[1] AND RCON1_EncodeOK[1] AND RCON1_IN[1].DataValid
       AND RCON1_MotionPermit[1] THEN
        E001_Out_OUT08_2003_09 := RCON1_TxUInt[8];
        E001_Out_OUT09_2003_0A := RCON1_TxUInt[9];
        E001_Out_OUT10_2003_0B := RCON1_TxUInt[10];
        E001_Out_OUT11_2003_0C := RCON1_TxUInt[11];
        E001_Out_OUT12_2003_0D := RCON1_TxUInt[12];
        E001_Out_OUT13_2003_0E := RCON1_TxUInt[13];
        E001_Out_OUT14_2003_0F := RCON1_TxUInt[14];
        E001_Out_OUT15_2003_10 := RCON1_TxUInt[15];
        RCON1_AxisWritten[1] := TRUE;
    END_IF;

// 2軸目＝実機軸No.1。OUT16～OUT23の8ワードをまとめて代入。
// AxisApply=この軸の更新許可、EncodeOK=変換OK、DataValid=入力情報の条件確認、MotionPermit=機械側の運転許可。
// 途中1ワードだけではなく、位置・幅・速度・加減速・押付け・制御を一組として渡します。
    IF RCON1_AxisApply[2] AND RCON1_EncodeOK[2] AND RCON1_IN[2].DataValid
       AND RCON1_MotionPermit[2] THEN
        E001_Out_OUT16_2003_11 := RCON1_TxUInt[16];
        E001_Out_OUT17_2003_12 := RCON1_TxUInt[17];
        E001_Out_OUT18_2003_13 := RCON1_TxUInt[18];
        E001_Out_OUT19_2003_14 := RCON1_TxUInt[19];
        E001_Out_OUT20_2003_15 := RCON1_TxUInt[20];
        E001_Out_OUT21_2003_16 := RCON1_TxUInt[21];
        E001_Out_OUT22_2003_17 := RCON1_TxUInt[22];
        E001_Out_OUT23_2003_18 := RCON1_TxUInt[23];
        RCON1_AxisWritten[2] := TRUE;
    END_IF;

// 3軸目＝実機軸No.2。OUT24～OUT31の8ワードをまとめて代入。
// AxisApply=この軸の更新許可、EncodeOK=変換OK、DataValid=入力情報の条件確認、MotionPermit=機械側の運転許可。
// 途中1ワードだけではなく、位置・幅・速度・加減速・押付け・制御を一組として渡します。
    IF RCON1_AxisApply[3] AND RCON1_EncodeOK[3] AND RCON1_IN[3].DataValid
       AND RCON1_MotionPermit[3] THEN
        E001_Out_OUT24_2003_19 := RCON1_TxUInt[24];
        E001_Out_OUT25_2003_1A := RCON1_TxUInt[25];
        E001_Out_OUT26_2003_1B := RCON1_TxUInt[26];
        E001_Out_OUT27_2003_1C := RCON1_TxUInt[27];
        E001_Out_OUT28_2003_1D := RCON1_TxUInt[28];
        E001_Out_OUT29_2003_1E := RCON1_TxUInt[29];
        E001_Out_OUT30_2003_1F := RCON1_TxUInt[30];
        E001_Out_OUT31_2003_20 := RCON1_TxUInt[31];
        RCON1_AxisWritten[3] := TRUE;
    END_IF;

// 4軸目＝実機軸No.3。OUT32～OUT39の8ワードをまとめて代入。
// AxisApply=この軸の更新許可、EncodeOK=変換OK、DataValid=入力情報の条件確認、MotionPermit=機械側の運転許可。
// 途中1ワードだけではなく、位置・幅・速度・加減速・押付け・制御を一組として渡します。
    IF RCON1_AxisApply[4] AND RCON1_EncodeOK[4] AND RCON1_IN[4].DataValid
       AND RCON1_MotionPermit[4] THEN
        E001_Out_OUT32_2003_21 := RCON1_TxUInt[32];
        E001_Out_OUT33_2003_22 := RCON1_TxUInt[33];
        E001_Out_OUT34_2003_23 := RCON1_TxUInt[34];
        E001_Out_OUT35_2003_24 := RCON1_TxUInt[35];
        E001_Out_OUT36_2003_25 := RCON1_TxUInt[36];
        E001_Out_OUT37_2003_26 := RCON1_TxUInt[37];
        E001_Out_OUT38_2003_27 := RCON1_TxUInt[38];
        E001_Out_OUT39_2003_28 := RCON1_TxUInt[39];
        RCON1_AxisWritten[4] := TRUE;
    END_IF;

// 5軸目＝実機軸No.4。OUT40～OUT47の8ワードをまとめて代入。
// AxisApply=この軸の更新許可、EncodeOK=変換OK、DataValid=入力情報の条件確認、MotionPermit=機械側の運転許可。
// 途中1ワードだけではなく、位置・幅・速度・加減速・押付け・制御を一組として渡します。
    IF RCON1_AxisApply[5] AND RCON1_EncodeOK[5] AND RCON1_IN[5].DataValid
       AND RCON1_MotionPermit[5] THEN
        E001_Out_OUT40_2003_29 := RCON1_TxUInt[40];
        E001_Out_OUT41_2003_2A := RCON1_TxUInt[41];
        E001_Out_OUT42_2003_2B := RCON1_TxUInt[42];
        E001_Out_OUT43_2003_2C := RCON1_TxUInt[43];
        E001_Out_OUT44_2003_2D := RCON1_TxUInt[44];
        E001_Out_OUT45_2003_2E := RCON1_TxUInt[45];
        E001_Out_OUT46_2003_2F := RCON1_TxUInt[46];
        E001_Out_OUT47_2003_30 := RCON1_TxUInt[47];
        RCON1_AxisWritten[5] := TRUE;
    END_IF;

// 6軸目＝実機軸No.5。OUT48～OUT55の8ワードをまとめて代入。
// AxisApply=この軸の更新許可、EncodeOK=変換OK、DataValid=入力情報の条件確認、MotionPermit=機械側の運転許可。
// 途中1ワードだけではなく、位置・幅・速度・加減速・押付け・制御を一組として渡します。
    IF RCON1_AxisApply[6] AND RCON1_EncodeOK[6] AND RCON1_IN[6].DataValid
       AND RCON1_MotionPermit[6] THEN
        E001_Out_OUT48_2003_31 := RCON1_TxUInt[48];
        E001_Out_OUT49_2003_32 := RCON1_TxUInt[49];
        E001_Out_OUT50_2003_33 := RCON1_TxUInt[50];
        E001_Out_OUT51_2003_34 := RCON1_TxUInt[51];
        E001_Out_OUT52_2003_35 := RCON1_TxUInt[52];
        E001_Out_OUT53_2003_36 := RCON1_TxUInt[53];
        E001_Out_OUT54_2003_37 := RCON1_TxUInt[54];
        E001_Out_OUT55_2003_38 := RCON1_TxUInt[55];
        RCON1_AxisWritten[6] := TRUE;
    END_IF;
END_IF;
// OUT01～07は予約領域のため書き換えません。OUT56以降は112Byte設定に存在しません。
// 現在の実機設定・別処理の用途が未確認なので、余剰領域を勝手にゼロクリアしません。
(* Rung 243: #RCON2/Node5 共通通信 / 入力変換 *)
// 【RCON2／Node5／5軸】直接数値指定の通信変換。加速と減速は共通値です。
// 前提：全軸が直接数値指定、直動軸、共通8ワード＋軸番号順に各8ワード。実機の設定は別途照合。
// OUTはPLC→RCONの指令、INはRCON→PLCの現在値・状態。名前はPLCから見た方向です。
// 構造体は人が扱いやすい箱、Eで始まる変数はI/Oマップに割付済みの通信の出入口です。
// このSTは変換と許可付き代入までです。自動運転、通信正常判定、安全停止、開始受付の管理は含みません。
// Sysmacでの全体再ビルドと実機照合は未実施です。このファイルだけで実機へ転送しないでください。
// 【① 入力を読む → 単位を戻す → 構造体INへ入れる】
// まず56個のUINTをRxRawへコピーします。ここでは実入力変数へ一切代入しません。
// 軸データはIN08～47。IN48～55は読みますが、用途を勝手に決めません。
// RxRawは通信のまま、RxWordは必要なら上下バイトを入れ替えた後の値です。
// 注意：確認前も数値・状態は仮に復元します。DataValid=FALSEの値で機械を動かさないでください。
RCON2_RxRaw[0] := E005_In_IN00_2004_01_1;
RCON2_RxRaw[1] := E005_In_IN01_2004_02_1;
RCON2_RxRaw[2] := E005_In_IN02_2004_03_1;
RCON2_RxRaw[3] := E005_In_IN03_2004_04_1;
RCON2_RxRaw[4] := E005_In_IN04_2004_05_1;
RCON2_RxRaw[5] := E005_In_IN05_2004_06_1;
RCON2_RxRaw[6] := E005_In_IN06_2004_07_1;
RCON2_RxRaw[7] := E005_In_IN07_2004_08_1;
RCON2_RxRaw[8] := E005_In_IN08_2004_09_1;
RCON2_RxRaw[9] := E005_In_IN09_2004_0A_1;
RCON2_RxRaw[10] := E005_In_IN10_2004_0B_1;
RCON2_RxRaw[11] := E005_In_IN11_2004_0C_1;
RCON2_RxRaw[12] := E005_In_IN12_2004_0D_1;
RCON2_RxRaw[13] := E005_In_IN13_2004_0E_1;
RCON2_RxRaw[14] := E005_In_IN14_2004_0F_1;
RCON2_RxRaw[15] := E005_In_IN15_2004_10_1;
RCON2_RxRaw[16] := E005_In_IN16_2004_11_1;
RCON2_RxRaw[17] := E005_In_IN17_2004_12_1;
RCON2_RxRaw[18] := E005_In_IN18_2004_13_1;
RCON2_RxRaw[19] := E005_In_IN19_2004_14_1;
RCON2_RxRaw[20] := E005_In_IN20_2004_15_1;
RCON2_RxRaw[21] := E005_In_IN21_2004_16_1;
RCON2_RxRaw[22] := E005_In_IN22_2004_17_1;
RCON2_RxRaw[23] := E005_In_IN23_2004_18_1;
RCON2_RxRaw[24] := E005_In_IN24_2004_19_1;
RCON2_RxRaw[25] := E005_In_IN25_2004_1A_1;
RCON2_RxRaw[26] := E005_In_IN26_2004_1B_1;
RCON2_RxRaw[27] := E005_In_IN27_2004_1C_1;
RCON2_RxRaw[28] := E005_In_IN28_2004_1D_1;
RCON2_RxRaw[29] := E005_In_IN29_2004_1E_1;
RCON2_RxRaw[30] := E005_In_IN30_2004_1F_1;
RCON2_RxRaw[31] := E005_In_IN31_2004_20_1;
RCON2_RxRaw[32] := E005_In_IN32_2004_21_1;
RCON2_RxRaw[33] := E005_In_IN33_2004_22_1;
RCON2_RxRaw[34] := E005_In_IN34_2004_23_1;
RCON2_RxRaw[35] := E005_In_IN35_2004_24_1;
RCON2_RxRaw[36] := E005_In_IN36_2004_25_1;
RCON2_RxRaw[37] := E005_In_IN37_2004_26_1;
RCON2_RxRaw[38] := E005_In_IN38_2004_27_1;
RCON2_RxRaw[39] := E005_In_IN39_2004_28_1;
RCON2_RxRaw[40] := E005_In_IN40_2004_29_1;
RCON2_RxRaw[41] := E005_In_IN41_2004_2A_1;
RCON2_RxRaw[42] := E005_In_IN42_2004_2B_1;
RCON2_RxRaw[43] := E005_In_IN43_2004_2C_1;
RCON2_RxRaw[44] := E005_In_IN44_2004_2D_1;
RCON2_RxRaw[45] := E005_In_IN45_2004_2E_1;
RCON2_RxRaw[46] := E005_In_IN46_2004_2F_1;
RCON2_RxRaw[47] := E005_In_IN47_2004_30_1;
RCON2_RxRaw[48] := E005_In_IN48_2004_31_1;
RCON2_RxRaw[49] := E005_In_IN49_2004_32_1;
RCON2_RxRaw[50] := E005_In_IN50_2004_33_1;
RCON2_RxRaw[51] := E005_In_IN51_2004_34_1;
RCON2_RxRaw[52] := E005_In_IN52_2004_35_1;
RCON2_RxRaw[53] := E005_In_IN53_2004_36_1;
RCON2_RxRaw[54] := E005_In_IN54_2004_37_1;
RCON2_RxRaw[55] := E005_In_IN55_2004_38_1;

// 取説の論理ワードへ正規化。Swapは1ワード内の上下バイト交換です。
// SwapBytesは推測で設定せず、既知の位置とbitで実機照合してください。
FOR ConvWordIndex := INT#0 TO INT#55 DO
    RCON2_RxWord[ConvWordIndex] := UINT_TO_WORD(RCON2_RxRaw[ConvWordIndex]);
    IF RCON2_SwapBytes THEN
        RCON2_RxWord[ConvWordIndex] := Swap(RCON2_RxWord[ConvWordIndex]);
    END_IF;
END_FOR;

ConvUnitOK := (RCON2_SpeedUnit_mm_s = LREAL#1.0) OR
              (RCON2_SpeedUnit_mm_s = LREAL#0.1);

// 【①-2 共通状態】IN00はユニット全体、IN01は各軸のリンク情報です。
// TestABit(ワード, bit番号)は、そのスイッチがONかをBOOLで取り出す命令です。
// 例：IN01のb0は軸No.0→配列[1]、b1は軸No.1→配列[2]。配列番号と実機軸番号は1違います。
// 共通固定領域。ここで使うbit番号は取説の論理bitです（MJ0384 6-24～6-25）。
RCON2_GwRun := TestABit(RCON2_RxWord[0], USINT#15);
RCON2_GwControllerCommLatch := TestABit(RCON2_RxWord[0], USINT#14);
RCON2_GwAxisCommError := TestABit(RCON2_RxWord[0], USINT#13);
RCON2_GwManual := TestABit(RCON2_RxWord[0], USINT#12);
RCON2_GwHeavyAlarm := TestABit(RCON2_RxWord[0], USINT#11);
RCON2_GwLightAlarm := TestABit(RCON2_RxWord[0], USINT#10);
RCON2_GwSystemStop := TestABit(RCON2_RxWord[0], USINT#8);
RCON2_GwAlarmCode := WORD_TO_UINT(RCON2_RxWord[0] AND WORD#16#00FF);
FOR ConvWordIndex := INT#0 TO INT#4 DO
    RCON2_PowerStateRaw[ConvWordIndex] := RCON2_RxWord[ConvWordIndex + INT#2];
END_FOR;

// 【①-3 軸ごとに同じ読取りを繰り返す】
// FORは1～5軸を順番に処理します。ConvBaseはその軸の先頭番号です。
// 計算：8+(軸番号-1)×8。1軸目=8、2軸目=16、3軸目=24。先頭8ワードは共通領域です。
FOR ConvAxisIndex := INT#1 TO INT#5 DO
    ConvBase := INT#8 + (ConvAxisIndex - INT#1) * INT#8;
    RCON2_AxisLinked[ConvAxisIndex] :=
        TestABit(RCON2_RxWord[1], INT_TO_USINT(ConvAxisIndex - INT#1));

// 例：下位2540／上位0なら32bit値2540→25.40mm。
// 上位を16bit左に動かして下位とORで重ねます。SHLが左シフト、ORがビットの合成です。
// 負位置はDWORD_TO_DINTで符号を復元。下位62996／上位65535なら-2540→-25.40mm。
    // 現在位置：下位・上位を結合、符号付き32bitとして解釈、0.01mmをmmへ。
    ConvDWord := SHL(WORD_TO_DWORD(RCON2_RxWord[ConvBase + INT#1]), ULINT#16)
                 OR WORD_TO_DWORD(RCON2_RxWord[ConvBase]);
    RCON2_IN[ConvAxisIndex].ActualPos_mm :=
        DINT_TO_LREAL(DWORD_TO_DINT(ConvDWord)) * LREAL#0.01;

    // 電流：32bitのmA。RCON-PCでは指令電流であり、実測トルクではありません。
    ConvDWord := SHL(WORD_TO_DWORD(RCON2_RxWord[ConvBase + INT#3]), ULINT#16)
                 OR WORD_TO_DWORD(RCON2_RxWord[ConvBase + INT#2]);
    RCON2_IN[ConvAxisIndex].Current_mA := DWORD_TO_DINT(ConvDWord);

    // 現在速度：16bitの負数をINTとして読む。UINTのまま速度にしません。
    IF ConvUnitOK THEN
        RCON2_IN[ConvAxisIndex].ActualSpeed_mm_s :=
            INT_TO_LREAL(WORD_TO_INT(RCON2_RxWord[ConvBase + INT#4])) * RCON2_SpeedUnit_mm_s;
    END_IF;
    // 単位不明のとき速度は前値を保持し、DataValidはFALSEにします。
    // 軸内の+5ワードは予約のため値を使用しません。
    RCON2_IN[ConvAxisIndex].AlarmCode := WORD_TO_UINT(RCON2_RxWord[ConvBase + INT#6]);

// 例：Status.ServoReady=TRUEは「サーボON状態を受信した」という意味。
// OUT側Control.ServoOn=TRUEは「サーボONを要求する」という意味で、指令と結果を区別します。
    // 状態ワード：12個のBOOLへ分解。予約b6,b9～11は使いません。
    RCON2_IN[ConvAxisIndex].Status.PositionDone := TestABit(RCON2_RxWord[ConvBase + INT#7], USINT#0);
    RCON2_IN[ConvAxisIndex].Status.HomeDone := TestABit(RCON2_RxWord[ConvBase + INT#7], USINT#1);
    RCON2_IN[ConvAxisIndex].Status.Moving := TestABit(RCON2_RxWord[ConvBase + INT#7], USINT#2);
    RCON2_IN[ConvAxisIndex].Status.Alarm := TestABit(RCON2_RxWord[ConvBase + INT#7], USINT#3);
    RCON2_IN[ConvAxisIndex].Status.ServoReady := TestABit(RCON2_RxWord[ConvBase + INT#7], USINT#4);
    RCON2_IN[ConvAxisIndex].Status.PushMiss := TestABit(RCON2_RxWord[ConvBase + INT#7], USINT#5);
    RCON2_IN[ConvAxisIndex].Status.OverloadWarning := TestABit(RCON2_RxWord[ConvBase + INT#7], USINT#7);
    RCON2_IN[ConvAxisIndex].Status.CommandDone := TestABit(RCON2_RxWord[ConvBase + INT#7], USINT#8);
    RCON2_IN[ConvAxisIndex].Status.Zone1 := TestABit(RCON2_RxWord[ConvBase + INT#7], USINT#12);
    RCON2_IN[ConvAxisIndex].Status.Zone2 := TestABit(RCON2_RxWord[ConvBase + INT#7], USINT#13);
    RCON2_IN[ConvAxisIndex].Status.ControllerReady := TestABit(RCON2_RxWord[ConvBase + INT#7], USINT#14);
    RCON2_IN[ConvAxisIndex].Status.EmergencyStop := TestABit(RCON2_RxWord[ConvBase + INT#7], USINT#15);

    // DataValidは直接受信bitではなく、今回の内部設計で決めた内部判定です。
    // CommOKはCPUの実通信状態から別途作成。単にTRUE固定にしないでください。
    // DataValidは運転許可や安全保証ではありません。各異常・原点等は別途確認。
    RCON2_IN[ConvAxisIndex].DataValid := RCON2_CommOK AND RCON2_LayoutConfirmed
        AND RCON2_ByteOrderConfirmed AND ConvUnitOK AND RCON2_GwRun
        AND RCON2_AxisLinked[ConvAxisIndex] AND NOT RCON2_GwAxisCommError;
END_FOR;

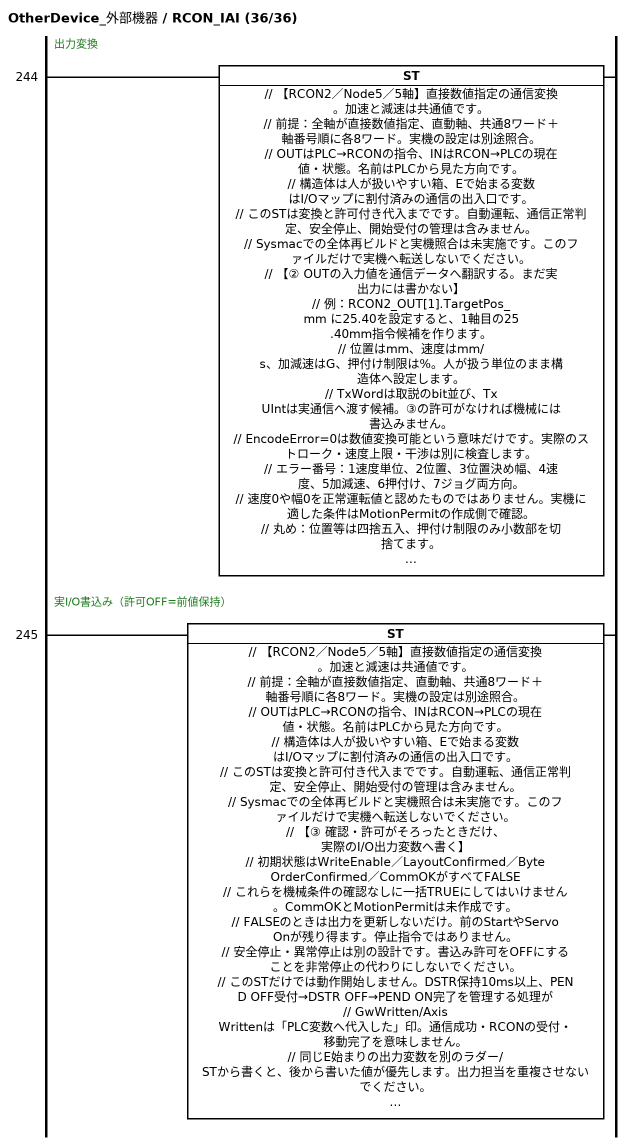
(* Rung 244: 出力変換 *)
// 【RCON2／Node5／5軸】直接数値指定の通信変換。加速と減速は共通値です。
// 前提：全軸が直接数値指定、直動軸、共通8ワード＋軸番号順に各8ワード。実機の設定は別途照合。
// OUTはPLC→RCONの指令、INはRCON→PLCの現在値・状態。名前はPLCから見た方向です。
// 構造体は人が扱いやすい箱、Eで始まる変数はI/Oマップに割付済みの通信の出入口です。
// このSTは変換と許可付き代入までです。自動運転、通信正常判定、安全停止、開始受付の管理は含みません。
// Sysmacでの全体再ビルドと実機照合は未実施です。このファイルだけで実機へ転送しないでください。
// 【② OUTの入力値を通信データへ翻訳する。まだ実出力には書かない】
// 例：RCON2_OUT[1].TargetPos_mm に25.40を設定すると、1軸目の25.40mm指令候補を作ります。
// 位置はmm、速度はmm/s、加減速はG、押付け制限は%。人が扱う単位のまま構造体へ設定します。
// TxWordは取説のbit並び、TxUIntは実通信へ渡す候補。③の許可がなければ機械には書込みません。
// EncodeError=0は数値変換可能という意味だけです。実際のストローク・速度上限・干渉は別に検査します。
// エラー番号：1速度単位、2位置、3位置決め幅、4速度、5加減速、6押付け、7ジョグ両方向。
// 速度0や幅0を正常運転値と認めたものではありません。実機に適した条件はMotionPermitの作成側で確認。
// 丸め：位置等は四捨五入、押付け制限のみ小数部を切捨てます。

ConvUnitOK := (RCON2_SpeedUnit_mm_s = LREAL#1.0) OR
              (RCON2_SpeedUnit_mm_s = LREAL#0.1);

// 共通制御：MONは論理b15、RTEは論理b13。他のbitは0。
// MONを落とす処理を安全停止として扱わないでください。
RCON2_TxWord[0] := WORD#16#0000;
IF RCON2_GwMON_Request THEN
    RCON2_TxWord[0] := RCON2_TxWord[0] OR WORD#16#8000;
END_IF;
IF RCON2_GwRTE_Request THEN
    RCON2_TxWord[0] := RCON2_TxWord[0] OR WORD#16#2000;
END_IF;

FOR ConvAxisIndex := INT#1 TO INT#5 DO
    ConvBase := INT#8 + (ConvAxisIndex - INT#1) * INT#8;
    RCON2_EncodeError[ConvAxisIndex] := UINT#0;

    // 比較で範囲を確認してから型変換するため、NaN・無限大も変換対象から外れます。
    // 位置・幅9999.99mmはこの案で採用する通信範囲の上限で、実機ストロークではありません。
    IF NOT ConvUnitOK THEN
        RCON2_EncodeError[ConvAxisIndex] := UINT#1;
    ELSIF NOT ((RCON2_OUT[ConvAxisIndex].TargetPos_mm >= LREAL#-9999.99) AND
               (RCON2_OUT[ConvAxisIndex].TargetPos_mm <= LREAL#9999.99)) THEN
        RCON2_EncodeError[ConvAxisIndex] := UINT#2;
    ELSIF NOT ((RCON2_OUT[ConvAxisIndex].PositionBand_mm >= LREAL#0.0) AND
               (RCON2_OUT[ConvAxisIndex].PositionBand_mm <= LREAL#9999.99)) THEN
        RCON2_EncodeError[ConvAxisIndex] := UINT#3;
    ELSIF NOT ((RCON2_OUT[ConvAxisIndex].Speed_mm_s >= LREAL#0.0) AND
               (RCON2_OUT[ConvAxisIndex].Speed_mm_s <= LREAL#65535.0 * RCON2_SpeedUnit_mm_s)) THEN
        RCON2_EncodeError[ConvAxisIndex] := UINT#4;
    ELSIF NOT ((RCON2_OUT[ConvAxisIndex].AccDec_G >= LREAL#0.0) AND
               (RCON2_OUT[ConvAxisIndex].AccDec_G <= LREAL#655.35)) THEN
        RCON2_EncodeError[ConvAxisIndex] := UINT#5;
    ELSIF NOT ((RCON2_OUT[ConvAxisIndex].PushLimit_pct >= LREAL#0.0) AND
               (RCON2_OUT[ConvAxisIndex].PushLimit_pct <= LREAL#200.0)) THEN
        RCON2_EncodeError[ConvAxisIndex] := UINT#6;
    ELSIF RCON2_OUT[ConvAxisIndex].Control.JogMinus AND RCON2_OUT[ConvAxisIndex].Control.JogPlus THEN
        RCON2_EncodeError[ConvAxisIndex] := UINT#7;
    END_IF;

    RCON2_EncodeOK[ConvAxisIndex] := RCON2_EncodeError[ConvAxisIndex] = UINT#0;
    IF RCON2_EncodeOK[ConvAxisIndex] THEN
    // 【数値例】TargetPos_mm=25.40→×100で2540。下位ワード2540、上位ワード0。
// 700.25mm→70025なので下位4489、上位1。65536を超えた分が上位に入ります。
// DINTは符号付きの数、DWORDは同じ32bitの模様。負数の符号を壊さず分割するために使い分けます。
// TRUNCは小数部を捨てます。正数+0.5／負数-0.5を先に行い、四捨五入を明示しています。
    // 目標位置：mmから0.01mmの符号付き整数へ。
        ConvScaled := RCON2_OUT[ConvAxisIndex].TargetPos_mm * LREAL#100.0;
        IF ConvScaled >= LREAL#0.0 THEN
            ConvPos := LINT_TO_DINT(TRUNC(ConvScaled + LREAL#0.5));
        ELSE
            ConvPos := LINT_TO_DINT(TRUNC(ConvScaled - LREAL#0.5));
        END_IF;
        // 負数を含む32bitパターンを保ち、下位・上位の16bitへ分割。
        ConvDWord := DINT_TO_DWORD(ConvPos);
        RCON2_TxWord[ConvBase] := DWORD_TO_WORD(ConvDWord AND DWORD#16#0000FFFF);
        RCON2_TxWord[ConvBase + INT#1] := DWORD_TO_WORD(SHR(ConvDWord, ULINT#16));

        // 位置決め幅：非負の内部整数としてUDINTを選定（メーカーの符号なし保証ではありません）。
        ConvBand := LINT_TO_UDINT(TRUNC(RCON2_OUT[ConvAxisIndex].PositionBand_mm * LREAL#100.0 + LREAL#0.5));
        ConvDWord := UDINT_TO_DWORD(ConvBand);
        RCON2_TxWord[ConvBase + INT#2] := DWORD_TO_WORD(ConvDWord AND DWORD#16#0000FFFF);
        RCON2_TxWord[ConvBase + INT#3] := DWORD_TO_WORD(SHR(ConvDWord, ULINT#16));

// 速度20mm/s：速度単位1.0なら20、0.1なら200を送信します。
// 加減速0.20G：×100して20。加速と減速の両方に同じ値を使います。
// 押付け50%：×255÷100=127.5を切捨てて127。押付けの使用可否・上限は実機仕様で別確認。
        // 速度は1カウント量が1.0か0.1かで値が10倍変わります。
        ConvSpeed := LINT_TO_UINT(TRUNC(RCON2_OUT[ConvAxisIndex].Speed_mm_s / RCON2_SpeedUnit_mm_s + LREAL#0.5));
        ConvAccDec := LINT_TO_UINT(TRUNC(RCON2_OUT[ConvAxisIndex].AccDec_G * LREAL#100.0 + LREAL#0.5));
        ConvPush := LINT_TO_UINT(TRUNC(RCON2_OUT[ConvAxisIndex].PushLimit_pct * LREAL#255.0 / LREAL#100.0));
        RCON2_TxWord[ConvBase + INT#4] := UINT_TO_WORD(ConvSpeed);
        RCON2_TxWord[ConvBase + INT#5] := UINT_TO_WORD(ConvAccDec);
        RCON2_TxWord[ConvBase + INT#6] := UINT_TO_WORD(ConvPush);
    END_IF;
    // 不正値の場合、数値ワードは前値保持。EncodeOK=FALSEで03の書込みを抑止。
    // 前値保持は停止指令ではありません。停止・異常処理は別途設計してください。

    // Controlを論理bitへ詰める。予約b9は必ず0。
    RCON2_TxWord[ConvBase + INT#7] := WORD#16#0000;
// b0 DSTR／Control.Start：TRUEで開始要求。受付応答と10ms以上の保持を確認してOFF。常時ONにしない。
    IF RCON2_OUT[ConvAxisIndex].Control.Start THEN
        RCON2_TxWord[ConvBase + INT#7] := RCON2_TxWord[ConvBase + INT#7] OR WORD#16#0001;
    END_IF;
// b1 HOME／Control.Home：TRUEで原点復帰を指令。原点復帰完了はIN側HomeDoneで確認。
    IF RCON2_OUT[ConvAxisIndex].Control.Home THEN
        RCON2_TxWord[ConvBase + INT#7] := RCON2_TxWord[ConvBase + INT#7] OR WORD#16#0002;
    END_IF;
// b2 STP／Control.Pause：TRUEで一時停止、FALSEで解除。非常停止・安全停止の代用ではない。
    IF RCON2_OUT[ConvAxisIndex].Control.Pause THEN
        RCON2_TxWord[ConvBase + INT#7] := RCON2_TxWord[ConvBase + INT#7] OR WORD#16#0004;
    END_IF;
// b3 RES／Control.Reset：TRUEでアラームリセット要求。コールドスタート級の異常には使用できない。
    IF RCON2_OUT[ConvAxisIndex].Control.Reset THEN
        RCON2_TxWord[ConvBase + INT#7] := RCON2_TxWord[ConvBase + INT#7] OR WORD#16#0008;
    END_IF;
// b4 SON／Control.ServoOn：TRUEでサーボON要求。ON状態はIN側ServoReadyで確認。
    IF RCON2_OUT[ConvAxisIndex].Control.ServoOn THEN
        RCON2_TxWord[ConvBase + INT#7] := RCON2_TxWord[ConvBase + INT#7] OR WORD#16#0010;
    END_IF;
// b5 JISL／Control.InchingSelect：TRUEは一定距離のインチング、FALSEは押している間のジョグ。
    IF RCON2_OUT[ConvAxisIndex].Control.InchingSelect THEN
        RCON2_TxWord[ConvBase + INT#7] := RCON2_TxWord[ConvBase + INT#7] OR WORD#16#0020;
    END_IF;
// b6 JVEL／Control.JogSpeedSelect：FALSEは速度No.26・距離No.48、TRUEは速度No.47または指令速度・距離No.49。
    IF RCON2_OUT[ConvAxisIndex].Control.JogSpeedSelect THEN
        RCON2_TxWord[ConvBase + INT#7] := RCON2_TxWord[ConvBase + INT#7] OR WORD#16#0040;
    END_IF;
// b7 JOG-／Control.JogMinus：TRUEで原点方向へジョグ。反対方向指令との同時ONを防ぐ。
    IF RCON2_OUT[ConvAxisIndex].Control.JogMinus THEN
        RCON2_TxWord[ConvBase + INT#7] := RCON2_TxWord[ConvBase + INT#7] OR WORD#16#0080;
    END_IF;
// b8 JOG+／Control.JogPlus：TRUEで反原点方向へジョグ。反対方向指令との同時ONを防ぐ。
    IF RCON2_OUT[ConvAxisIndex].Control.JogPlus THEN
        RCON2_TxWord[ConvBase + INT#7] := RCON2_TxWord[ConvBase + INT#7] OR WORD#16#0100;
    END_IF;
// b10 GSL0／Control.GainSelect0：GainSelect1と組合せてサーボゲインセット0～3を選ぶ。機械調整用。
    IF RCON2_OUT[ConvAxisIndex].Control.GainSelect0 THEN
        RCON2_TxWord[ConvBase + INT#7] := RCON2_TxWord[ConvBase + INT#7] OR WORD#16#0400;
    END_IF;
// b11 GSL1／Control.GainSelect1：GainSelect0との2bitで選択。速度指令とは別の機能。
    IF RCON2_OUT[ConvAxisIndex].Control.GainSelect1 THEN
        RCON2_TxWord[ConvBase + INT#7] := RCON2_TxWord[ConvBase + INT#7] OR WORD#16#0800;
    END_IF;
// b12 PUSH／Control.PushEnable：TRUEは押付け、FALSEは通常位置決め。押付け条件は別途確認。
    IF RCON2_OUT[ConvAxisIndex].Control.PushEnable THEN
        RCON2_TxWord[ConvBase + INT#7] := RCON2_TxWord[ConvBase + INT#7] OR WORD#16#1000;
    END_IF;
// b13 DIR／Control.PushDirection：CON方式押付け時、TRUEは反原点方向、FALSEは原点方向。
    IF RCON2_OUT[ConvAxisIndex].Control.PushDirection THEN
        RCON2_TxWord[ConvBase + INT#7] := RCON2_TxWord[ConvBase + INT#7] OR WORD#16#2000;
    END_IF;
// b14 INC／Control.RelativeMove：FALSEは絶対座標、TRUEは現在位置からの相対移動量。
    IF RCON2_OUT[ConvAxisIndex].Control.RelativeMove THEN
        RCON2_TxWord[ConvBase + INT#7] := RCON2_TxWord[ConvBase + INT#7] OR WORD#16#4000;
    END_IF;
// b15 BKRL／Control.BrakeRelease：TRUEはブレーキ強制解除。通常FALSE。縦軸では落下等の危険がある。
    IF RCON2_OUT[ConvAxisIndex].Control.BrakeRelease THEN
        RCON2_TxWord[ConvBase + INT#7] := RCON2_TxWord[ConvBase + INT#7] OR WORD#16#8000;
    END_IF;
END_FOR;

// 論理ワードから実際に送るUINTへ。INと同じ1ワード内のバイト交換を適用します。
FOR ConvWordIndex := INT#0 TO INT#47 DO
    ConvWord := RCON2_TxWord[ConvWordIndex];
    IF RCON2_SwapBytes THEN
        ConvWord := Swap(ConvWord);
    END_IF;
    RCON2_TxUInt[ConvWordIndex] := WORD_TO_UINT(ConvWord);
END_FOR;
(* Rung 245: 実I/O書込み（許可OFF=前値保持） *)
// 【RCON2／Node5／5軸】直接数値指定の通信変換。加速と減速は共通値です。
// 前提：全軸が直接数値指定、直動軸、共通8ワード＋軸番号順に各8ワード。実機の設定は別途照合。
// OUTはPLC→RCONの指令、INはRCON→PLCの現在値・状態。名前はPLCから見た方向です。
// 構造体は人が扱いやすい箱、Eで始まる変数はI/Oマップに割付済みの通信の出入口です。
// このSTは変換と許可付き代入までです。自動運転、通信正常判定、安全停止、開始受付の管理は含みません。
// Sysmacでの全体再ビルドと実機照合は未実施です。このファイルだけで実機へ転送しないでください。
// 【③ 確認・許可がそろったときだけ、実際のI/O出力変数へ書く】
// 初期状態はWriteEnable／LayoutConfirmed／ByteOrderConfirmed／CommOKがすべてFALSEです。
// これらを機械条件の確認なしに一括TRUEにしてはいけません。CommOKとMotionPermitは未作成です。
// FALSEのときは出力を更新しないだけ。前のStartやServoOnが残り得ます。停止指令ではありません。
// 安全停止・異常停止は別の設計です。書込み許可をOFFにすることを非常停止の代わりにしないでください。
// このSTだけでは動作開始しません。DSTR保持10ms以上、PEND OFF受付→DSTR OFF→PEND ON完了を管理する処理が必要です。
// GwWritten/AxisWrittenは「PLC変数へ代入した」印。通信成功・RCONの受付・移動完了を意味しません。
// 同じE始まりの出力変数を別のラダー/STから書くと、後から書いた値が優先します。出力担当を重複させないでください。

RCON2_GwWritten := FALSE;
FOR ConvAxisIndex := INT#1 TO INT#5 DO
    RCON2_AxisWritten[ConvAxisIndex] := FALSE;
END_FOR;

IF RCON2_WriteEnable AND RCON2_LayoutConfirmed AND RCON2_ByteOrderConfirmed AND RCON2_CommOK THEN
// 共通指令はMON/RTEのみ。最初のRUN応答に必要なため、軸DataValidとは別にGwApplyで許可します。
    IF RCON2_GwApply THEN
        E005_Out_OUT00_2003_01_1 := RCON2_TxUInt[0];
        RCON2_GwWritten := TRUE;
    END_IF;

// 1軸目＝実機軸No.0。OUT08～OUT15の8ワードをまとめて代入。
// AxisApply=この軸の更新許可、EncodeOK=変換OK、DataValid=入力情報の条件確認、MotionPermit=機械側の運転許可。
// 途中1ワードだけではなく、位置・幅・速度・加減速・押付け・制御を一組として渡します。
    IF RCON2_AxisApply[1] AND RCON2_EncodeOK[1] AND RCON2_IN[1].DataValid
       AND RCON2_MotionPermit[1] THEN
        E005_Out_OUT08_2003_09_1 := RCON2_TxUInt[8];
        E005_Out_OUT09_2003_0A_1 := RCON2_TxUInt[9];
        E005_Out_OUT10_2003_0B_1 := RCON2_TxUInt[10];
        E005_Out_OUT11_2003_0C_1 := RCON2_TxUInt[11];
        E005_Out_OUT12_2003_0D_1 := RCON2_TxUInt[12];
        E005_Out_OUT13_2003_0E_1 := RCON2_TxUInt[13];
        E005_Out_OUT14_2003_0F_1 := RCON2_TxUInt[14];
        E005_Out_OUT15_2003_10_1 := RCON2_TxUInt[15];
        RCON2_AxisWritten[1] := TRUE;
    END_IF;

// 2軸目＝実機軸No.1。OUT16～OUT23の8ワードをまとめて代入。
// AxisApply=この軸の更新許可、EncodeOK=変換OK、DataValid=入力情報の条件確認、MotionPermit=機械側の運転許可。
// 途中1ワードだけではなく、位置・幅・速度・加減速・押付け・制御を一組として渡します。
    IF RCON2_AxisApply[2] AND RCON2_EncodeOK[2] AND RCON2_IN[2].DataValid
       AND RCON2_MotionPermit[2] THEN
        E005_Out_OUT16_2003_11_1 := RCON2_TxUInt[16];
        E005_Out_OUT17_2003_12_1 := RCON2_TxUInt[17];
        E005_Out_OUT18_2003_13_1 := RCON2_TxUInt[18];
        E005_Out_OUT19_2003_14_1 := RCON2_TxUInt[19];
        E005_Out_OUT20_2003_15_1 := RCON2_TxUInt[20];
        E005_Out_OUT21_2003_16_1 := RCON2_TxUInt[21];
        E005_Out_OUT22_2003_17_1 := RCON2_TxUInt[22];
        E005_Out_OUT23_2003_18_1 := RCON2_TxUInt[23];
        RCON2_AxisWritten[2] := TRUE;
    END_IF;

// 3軸目＝実機軸No.2。OUT24～OUT31の8ワードをまとめて代入。
// AxisApply=この軸の更新許可、EncodeOK=変換OK、DataValid=入力情報の条件確認、MotionPermit=機械側の運転許可。
// 途中1ワードだけではなく、位置・幅・速度・加減速・押付け・制御を一組として渡します。
    IF RCON2_AxisApply[3] AND RCON2_EncodeOK[3] AND RCON2_IN[3].DataValid
       AND RCON2_MotionPermit[3] THEN
        E005_Out_OUT24_2003_19_1 := RCON2_TxUInt[24];
        E005_Out_OUT25_2003_1A_1 := RCON2_TxUInt[25];
        E005_Out_OUT26_2003_1B_1 := RCON2_TxUInt[26];
        E005_Out_OUT27_2003_1C_1 := RCON2_TxUInt[27];
        E005_Out_OUT28_2003_1D_1 := RCON2_TxUInt[28];
        E005_Out_OUT29_2003_1E_1 := RCON2_TxUInt[29];
        E005_Out_OUT30_2003_1F_1 := RCON2_TxUInt[30];
        E005_Out_OUT31_2003_20_1 := RCON2_TxUInt[31];
        RCON2_AxisWritten[3] := TRUE;
    END_IF;

// 4軸目＝実機軸No.3。OUT32～OUT39の8ワードをまとめて代入。
// AxisApply=この軸の更新許可、EncodeOK=変換OK、DataValid=入力情報の条件確認、MotionPermit=機械側の運転許可。
// 途中1ワードだけではなく、位置・幅・速度・加減速・押付け・制御を一組として渡します。
    IF RCON2_AxisApply[4] AND RCON2_EncodeOK[4] AND RCON2_IN[4].DataValid
       AND RCON2_MotionPermit[4] THEN
        E005_Out_OUT32_2003_21_1 := RCON2_TxUInt[32];
        E005_Out_OUT33_2003_22_1 := RCON2_TxUInt[33];
        E005_Out_OUT34_2003_23_1 := RCON2_TxUInt[34];
        E005_Out_OUT35_2003_24_1 := RCON2_TxUInt[35];
        E005_Out_OUT36_2003_25_1 := RCON2_TxUInt[36];
        E005_Out_OUT37_2003_26_1 := RCON2_TxUInt[37];
        E005_Out_OUT38_2003_27_1 := RCON2_TxUInt[38];
        E005_Out_OUT39_2003_28_1 := RCON2_TxUInt[39];
        RCON2_AxisWritten[4] := TRUE;
    END_IF;

// 5軸目＝実機軸No.4。OUT40～OUT47の8ワードをまとめて代入。
// AxisApply=この軸の更新許可、EncodeOK=変換OK、DataValid=入力情報の条件確認、MotionPermit=機械側の運転許可。
// 途中1ワードだけではなく、位置・幅・速度・加減速・押付け・制御を一組として渡します。
    IF RCON2_AxisApply[5] AND RCON2_EncodeOK[5] AND RCON2_IN[5].DataValid
       AND RCON2_MotionPermit[5] THEN
        E005_Out_OUT40_2003_29_1 := RCON2_TxUInt[40];
        E005_Out_OUT41_2003_2A_1 := RCON2_TxUInt[41];
        E005_Out_OUT42_2003_2B_1 := RCON2_TxUInt[42];
        E005_Out_OUT43_2003_2C_1 := RCON2_TxUInt[43];
        E005_Out_OUT44_2003_2D_1 := RCON2_TxUInt[44];
        E005_Out_OUT45_2003_2E_1 := RCON2_TxUInt[45];
        E005_Out_OUT46_2003_2F_1 := RCON2_TxUInt[46];
        E005_Out_OUT47_2003_30_1 := RCON2_TxUInt[47];
        RCON2_AxisWritten[5] := TRUE;
    END_IF;
END_IF;
// OUT01～07、OUT48～55は、このSTからは一切書き換えません。
// 現在の実機設定・別処理の用途が未確認なので、余剰領域を勝手にゼロクリアしません。

(* Section DLEP1_GT2: ladder, written here as Structured Text *)

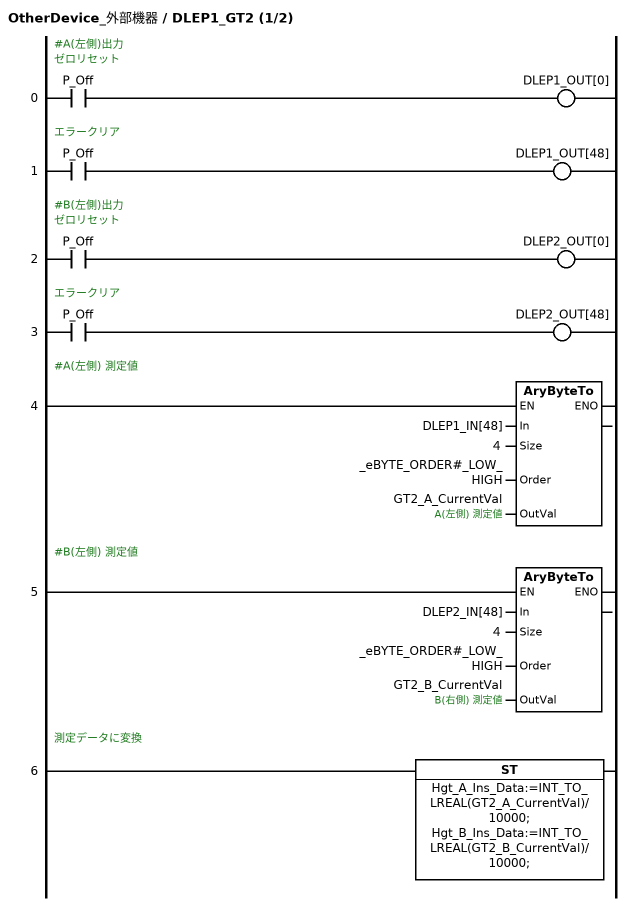
(* Rung 0: #A(左側)出力 / ゼロリセット *)
DLEP1_OUT[0] := P_Off;
(* Rung 1: エラークリア *)
DLEP1_OUT[48] := P_Off;
(* Rung 2: #B(左側)出力 / ゼロリセット *)
DLEP2_OUT[0] := P_Off;
(* Rung 3: エラークリア *)
DLEP2_OUT[48] := P_Off;
(* Rung 4: #A(左側) 測定値 *)
AryByteTo(In := DLEP1_IN[48], Size := ４, Order := _eBYTE_ORDER#_LOW_HIGH, OutVal := GT2_A_CurrentVal);
(* Rung 5: #B(左側) 測定値 *)
AryByteTo(In := DLEP2_IN[48], Size := ４, Order := _eBYTE_ORDER#_LOW_HIGH, OutVal := GT2_B_CurrentVal);
(* Rung 6: 測定データに変換 *)
Hgt_A_Ins_Data:=INT_TO_LREAL(GT2_A_CurrentVal)/10000;
Hgt_B_Ins_Data:=INT_TO_LREAL(GT2_B_CurrentVal)/10000;

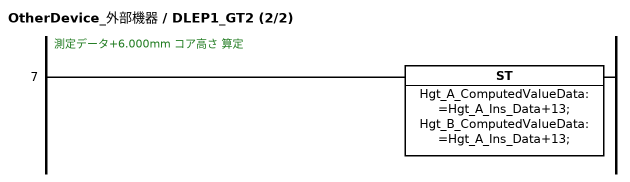
(* Rung 7: 測定データ+6.000mm コア高さ 算定 *)
Hgt_A_ComputedValueData:=Hgt_A_Ins_Data+13;
Hgt_B_ComputedValueData:=Hgt_A_Ins_Data+13;

(* Section FH_5552_10: ladder, written here as Structured Text *)

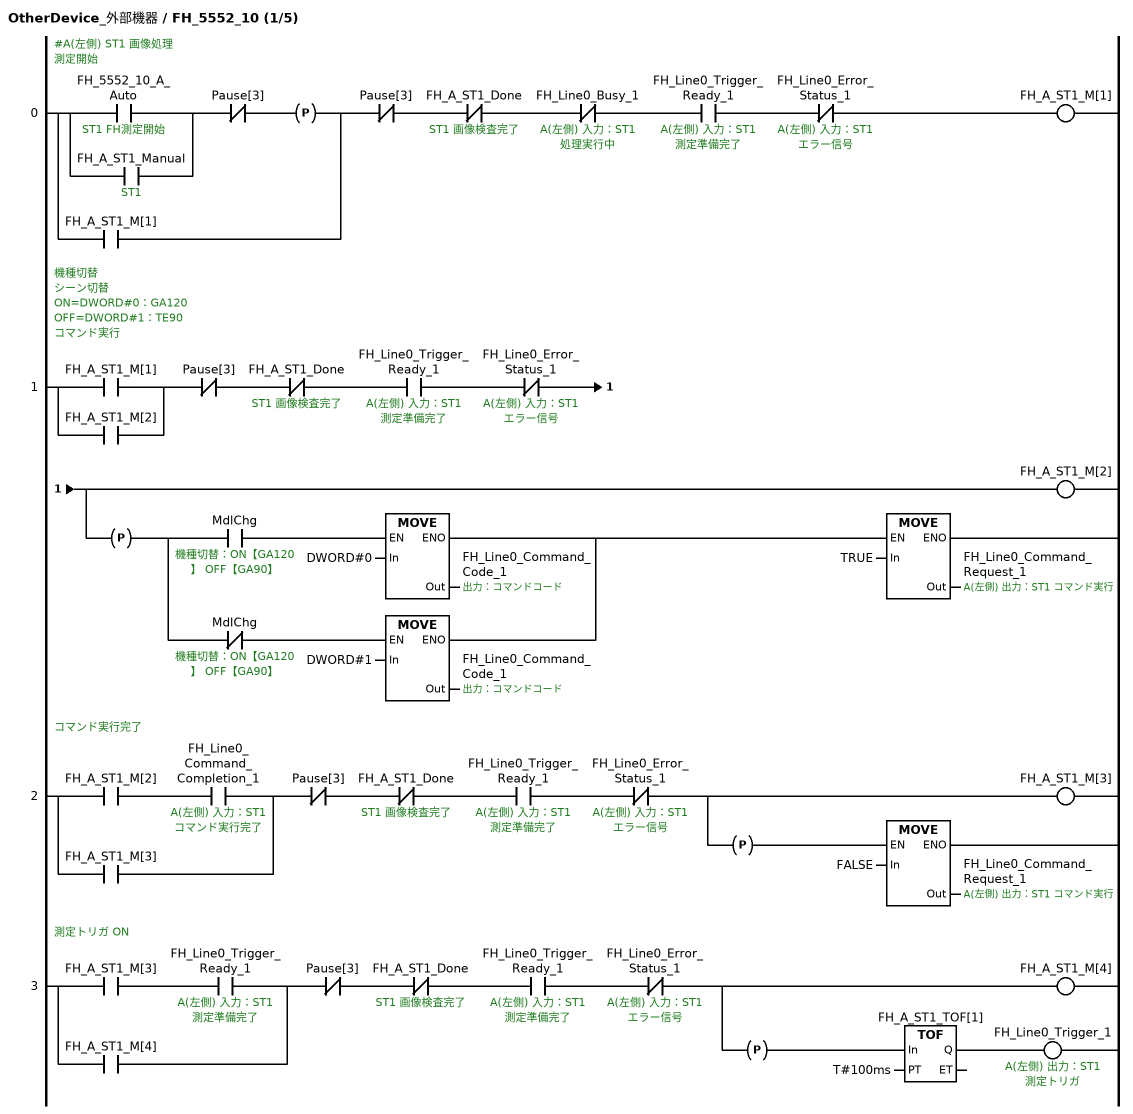
(* Rung 0: #A(左側) ST1 画像処理 / 測定開始 *)
_e25(CLK := (FH_5552_10_A_Auto OR FH_A_ST1_Manual) AND NOT Pause[3]);
FH_A_ST1_M[1] := (_e25.Q OR FH_A_ST1_M[1]) AND NOT Pause[3] AND NOT FH_A_ST1_Done AND NOT FH_Line0_Busy_1 AND FH_Line0_Trigger_Ready_1 AND NOT FH_Line0_Error_Status_1;
(* Rung 1: 機種切替 / シーン切替 / ON=DWORD#0：GA120 / OFF=DWORD#1：TE90 / コマンド実行 *)
_p26 := (FH_A_ST1_M[1] OR FH_A_ST1_M[2]) AND NOT Pause[3] AND NOT FH_A_ST1_Done AND FH_Line0_Trigger_Ready_1 AND NOT FH_Line0_Error_Status_1;
FH_A_ST1_M[2] := _p26;
_e27(CLK := _p26);
IF _e27.Q AND MdlChg THEN FH_Line0_Command_Code_1 := DWORD#0; END_IF;
IF _e27.Q AND NOT MdlChg THEN FH_Line0_Command_Code_1 := DWORD#1; END_IF;
IF _e27.Q AND (MdlChg OR NOT MdlChg) THEN FH_Line0_Command_Request_1 := TRUE; END_IF;
(* Rung 2: コマンド実行完了 *)
_p28 := ((FH_A_ST1_M[2] AND FH_Line0_Command_Completion_1) OR FH_A_ST1_M[3]) AND NOT Pause[3] AND NOT FH_A_ST1_Done AND FH_Line0_Trigger_Ready_1 AND NOT FH_Line0_Error_Status_1;
FH_A_ST1_M[3] := _p28;
_e29(CLK := _p28);
IF _e29.Q THEN FH_Line0_Command_Request_1 := FALSE; END_IF;
(* Rung 3: 測定トリガ ON *)
_p30 := ((FH_A_ST1_M[3] AND FH_Line0_Trigger_Ready_1) OR FH_A_ST1_M[4]) AND NOT Pause[3] AND NOT FH_A_ST1_Done AND FH_Line0_Trigger_Ready_1 AND NOT FH_Line0_Error_Status_1;
FH_A_ST1_M[4] := _p30;
_e31(CLK := _p30);
FH_A_ST1_TOF[1](In := _e31.Q, PT := T#100ms);
FH_Line0_Trigger_1 := FH_A_ST1_TOF[1].Q;

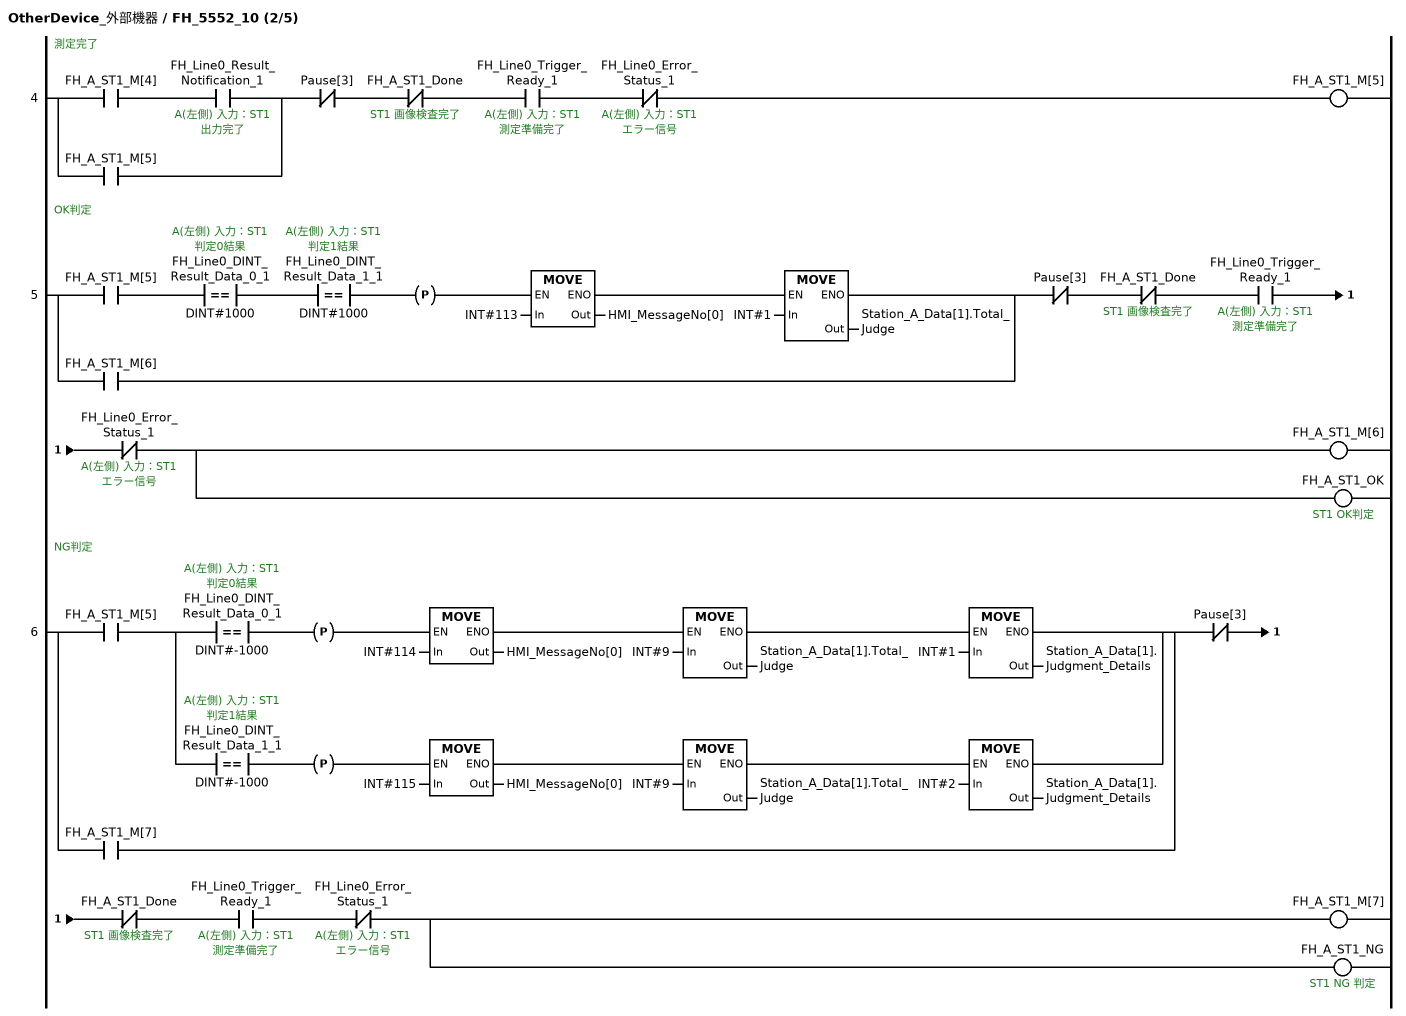
(* Rung 4: 測定完了 *)
FH_A_ST1_M[5] := ((FH_A_ST1_M[4] AND FH_Line0_Result_Notification_1) OR FH_A_ST1_M[5]) AND NOT Pause[3] AND NOT FH_A_ST1_Done AND FH_Line0_Trigger_Ready_1 AND NOT FH_Line0_Error_Status_1;
(* Rung 5: OK判定 *)
_e32(CLK := FH_A_ST1_M[5] AND (FH_Line0_DINT_Result_Data_0_1 = DINT#1000) AND (FH_Line0_DINT_Result_Data_1_1 = DINT#1000));
IF _e32.Q THEN
    HMI_MessageNo[0] := INT#113;
    Station_A_Data[1].Total_Judge := INT#1;
END_IF;
_p33 := (_e32.Q OR FH_A_ST1_M[6]) AND NOT Pause[3] AND NOT FH_A_ST1_Done AND FH_Line0_Trigger_Ready_1 AND NOT FH_Line0_Error_Status_1;
FH_A_ST1_M[6] := _p33;
FH_A_ST1_OK := _p33;
(* Rung 6: NG判定 *)
_e34(CLK := FH_A_ST1_M[5] AND (FH_Line0_DINT_Result_Data_0_1 = (DINT#-1000)));
IF _e34.Q THEN
    HMI_MessageNo[0] := INT#114;
    Station_A_Data[1].Total_Judge := INT#9;
    Station_A_Data[1].Judgment_Details := INT#1;
END_IF;
_e35(CLK := FH_A_ST1_M[5] AND (FH_Line0_DINT_Result_Data_1_1 = (DINT#-1000)));
IF _e35.Q THEN
    HMI_MessageNo[0] := INT#115;
    Station_A_Data[1].Total_Judge := INT#9;
    Station_A_Data[1].Judgment_Details := INT#2;
END_IF;
_p36 := (_e34.Q OR _e35.Q OR FH_A_ST1_M[7]) AND NOT Pause[3] AND NOT FH_A_ST1_Done AND FH_Line0_Trigger_Ready_1 AND NOT FH_Line0_Error_Status_1;
FH_A_ST1_M[7] := _p36;
FH_A_ST1_NG := _p36;

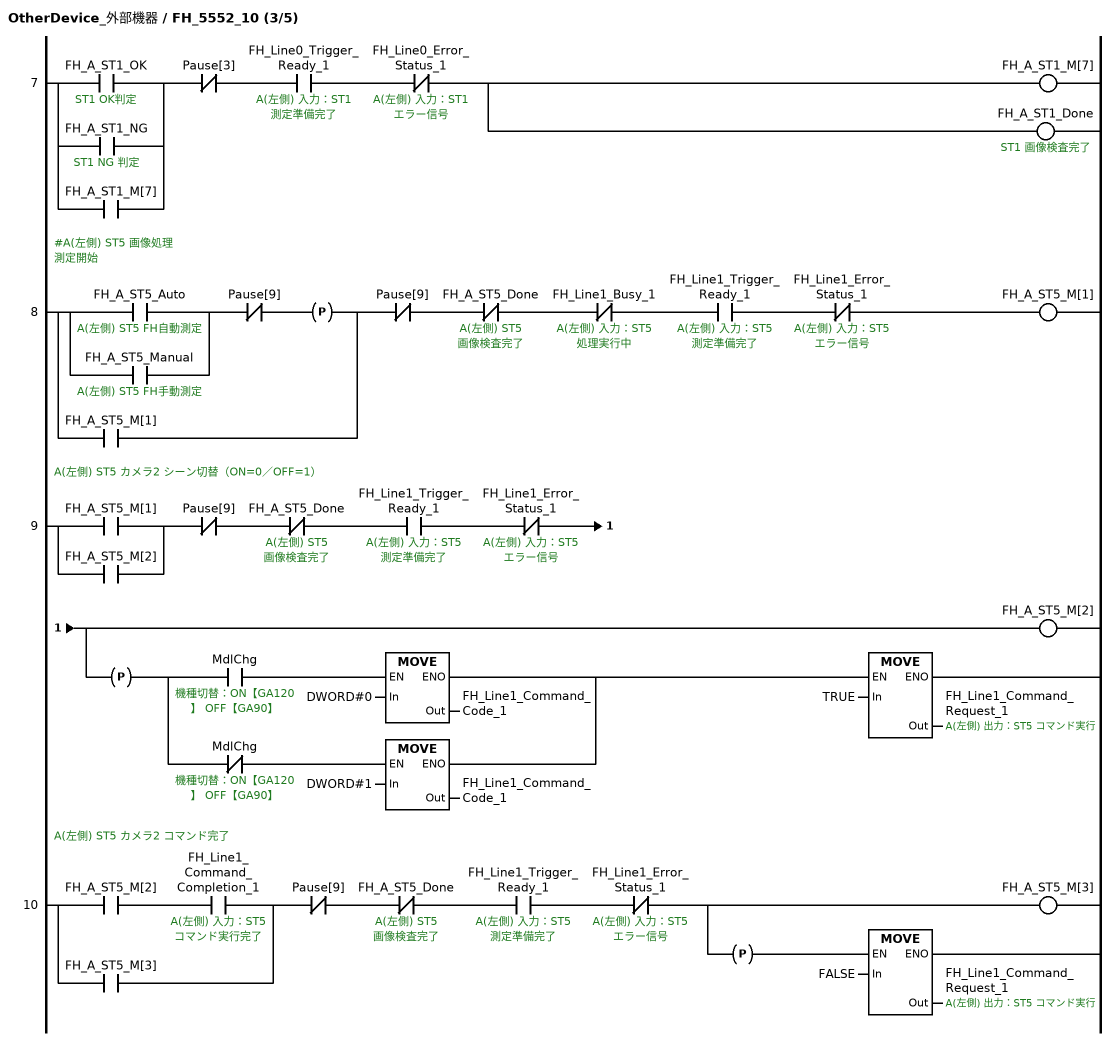
(* Rung 7 *)
_p37 := (FH_A_ST1_OK OR FH_A_ST1_NG OR FH_A_ST1_M[7]) AND NOT Pause[3] AND FH_Line0_Trigger_Ready_1 AND NOT FH_Line0_Error_Status_1;
FH_A_ST1_M[7] := _p37;
FH_A_ST1_Done := _p37;
(* Rung 8: #A(左側) ST5 画像処理 / 測定開始 *)
_e38(CLK := (FH_A_ST5_Auto OR FH_A_ST5_Manual) AND NOT Pause[9]);
FH_A_ST5_M[1] := (_e38.Q OR FH_A_ST5_M[1]) AND NOT Pause[9] AND NOT FH_A_ST5_Done AND NOT FH_Line1_Busy_1 AND FH_Line1_Trigger_Ready_1 AND NOT FH_Line1_Error_Status_1;
(* Rung 9: A(左側) ST5 カメラ2 シーン切替（ON=0／OFF=1） *)
_p39 := (FH_A_ST5_M[1] OR FH_A_ST5_M[2]) AND NOT Pause[9] AND NOT FH_A_ST5_Done AND FH_Line1_Trigger_Ready_1 AND NOT FH_Line1_Error_Status_1;
FH_A_ST5_M[2] := _p39;
_e40(CLK := _p39);
IF _e40.Q AND MdlChg THEN FH_Line1_Command_Code_1 := DWORD#0; END_IF;
IF _e40.Q AND NOT MdlChg THEN FH_Line1_Command_Code_1 := DWORD#1; END_IF;
IF _e40.Q AND (MdlChg OR NOT MdlChg) THEN FH_Line1_Command_Request_1 := TRUE; END_IF;
(* Rung 10: A(左側) ST5 カメラ2 コマンド完了 *)
_p41 := ((FH_A_ST5_M[2] AND FH_Line1_Command_Completion_1) OR FH_A_ST5_M[3]) AND NOT Pause[9] AND NOT FH_A_ST5_Done AND FH_Line1_Trigger_Ready_1 AND NOT FH_Line1_Error_Status_1;
FH_A_ST5_M[3] := _p41;
_e42(CLK := _p41);
IF _e42.Q THEN FH_Line1_Command_Request_1 := FALSE; END_IF;

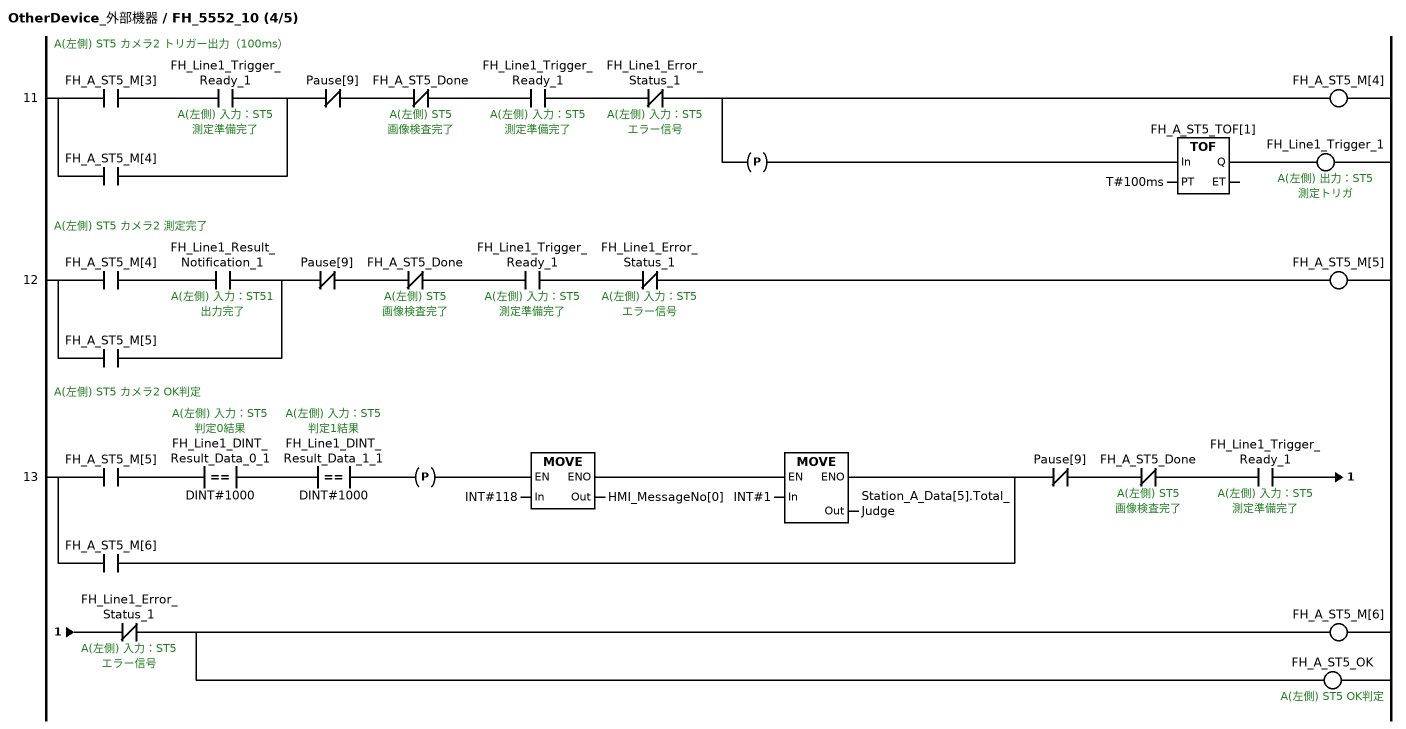
(* Rung 11: A(左側) ST5 カメラ2 トリガー出力（100ms） *)
_p43 := ((FH_A_ST5_M[3] AND FH_Line1_Trigger_Ready_1) OR FH_A_ST5_M[4]) AND NOT Pause[9] AND NOT FH_A_ST5_Done AND FH_Line1_Trigger_Ready_1 AND NOT FH_Line1_Error_Status_1;
FH_A_ST5_M[4] := _p43;
_e44(CLK := _p43);
FH_A_ST5_TOF[1](In := _e44.Q, PT := T#100ms);
FH_Line1_Trigger_1 := FH_A_ST5_TOF[1].Q;
(* Rung 12: A(左側) ST5 カメラ2 測定完了 *)
FH_A_ST5_M[5] := ((FH_A_ST5_M[4] AND FH_Line1_Result_Notification_1) OR FH_A_ST5_M[5]) AND NOT Pause[9] AND NOT FH_A_ST5_Done AND FH_Line1_Trigger_Ready_1 AND NOT FH_Line1_Error_Status_1;
(* Rung 13: A(左側) ST5 カメラ2 OK判定 *)
_e45(CLK := FH_A_ST5_M[5] AND (FH_Line1_DINT_Result_Data_0_1 = DINT#1000) AND (FH_Line1_DINT_Result_Data_1_1 = DINT#1000));
IF _e45.Q THEN
    HMI_MessageNo[0] := INT#118;
    Station_A_Data[5].Total_Judge := INT#1;
END_IF;
_p46 := (_e45.Q OR FH_A_ST5_M[6]) AND NOT Pause[9] AND NOT FH_A_ST5_Done AND FH_Line1_Trigger_Ready_1 AND NOT FH_Line1_Error_Status_1;
FH_A_ST5_M[6] := _p46;
FH_A_ST5_OK := _p46;

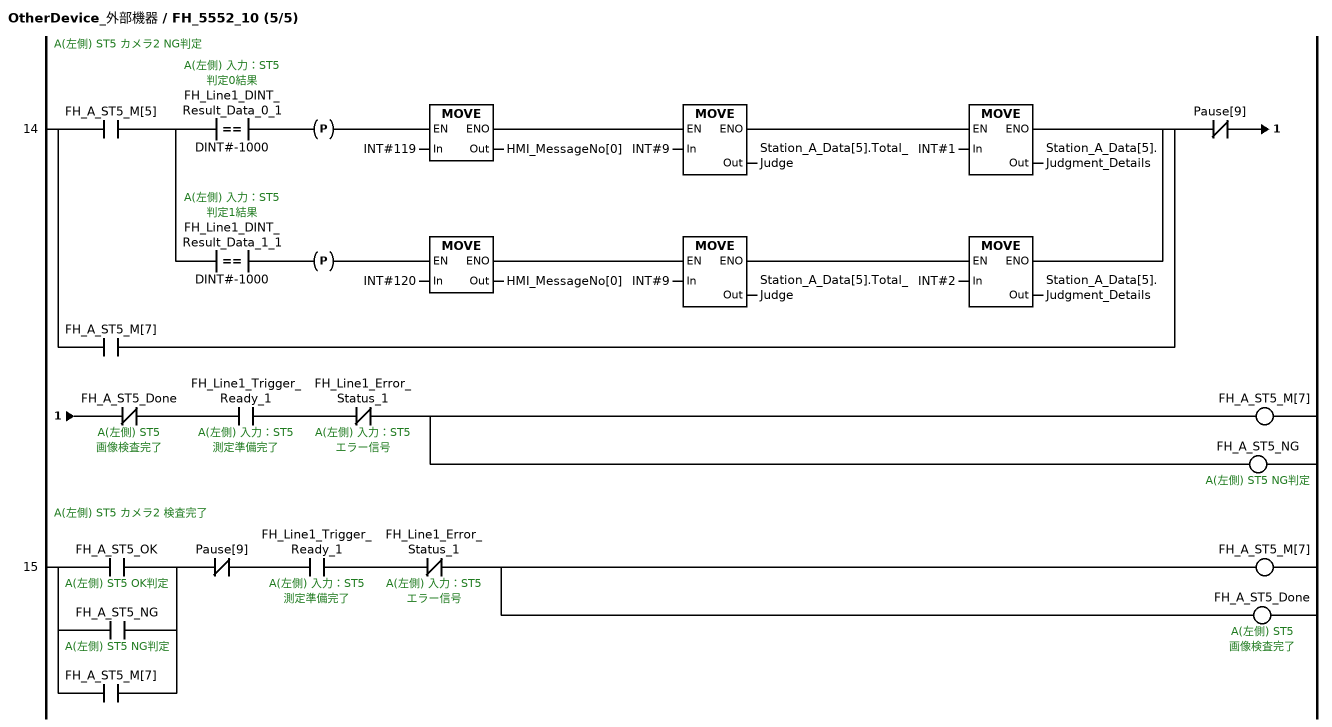
(* Rung 14: A(左側) ST5 カメラ2 NG判定 *)
_e47(CLK := FH_A_ST5_M[5] AND (FH_Line1_DINT_Result_Data_0_1 = (DINT#-1000)));
IF _e47.Q THEN
    HMI_MessageNo[0] := INT#119;
    Station_A_Data[5].Total_Judge := INT#9;
    Station_A_Data[5].Judgment_Details := INT#1;
END_IF;
_e48(CLK := FH_A_ST5_M[5] AND (FH_Line1_DINT_Result_Data_1_1 = (DINT#-1000)));
IF _e48.Q THEN
    HMI_MessageNo[0] := INT#120;
    Station_A_Data[5].Total_Judge := INT#9;
    Station_A_Data[5].Judgment_Details := INT#2;
END_IF;
_p49 := (_e47.Q OR _e48.Q OR FH_A_ST5_M[7]) AND NOT Pause[9] AND NOT FH_A_ST5_Done AND FH_Line1_Trigger_Ready_1 AND NOT FH_Line1_Error_Status_1;
FH_A_ST5_M[7] := _p49;
FH_A_ST5_NG := _p49;
(* Rung 15: A(左側) ST5 カメラ2 検査完了 *)
_p50 := (FH_A_ST5_OK OR FH_A_ST5_NG OR FH_A_ST5_M[7]) AND NOT Pause[9] AND FH_Line1_Trigger_Ready_1 AND NOT FH_Line1_Error_Status_1;
FH_A_ST5_M[7] := _p50;
FH_A_ST5_Done := _p50;

(* Section CV2A_KED: ladder, written here as Structured Text *)

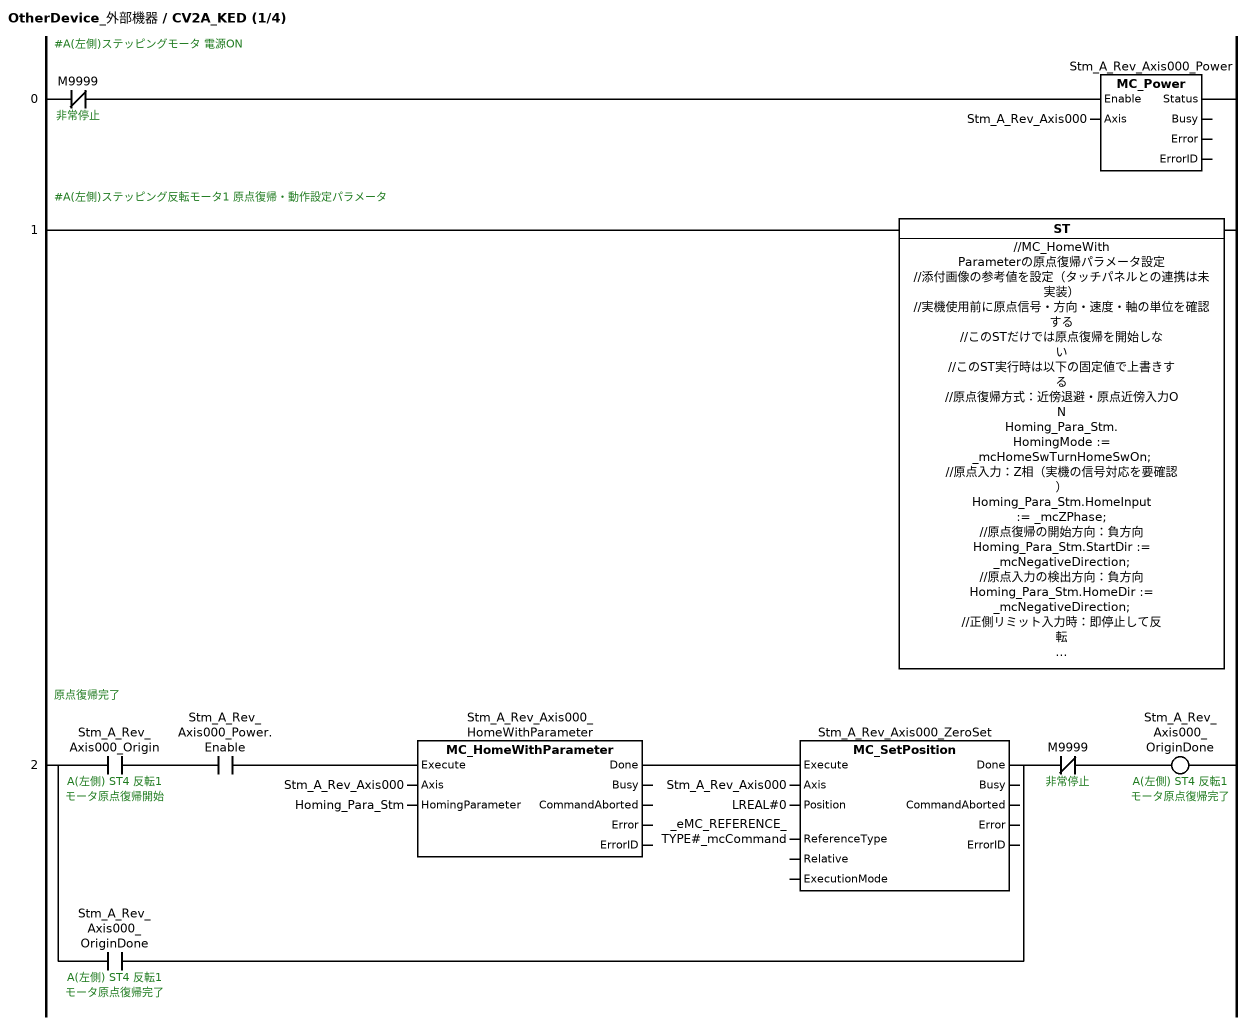
(* Rung 0: #A(左側)ステッピングモータ 電源ON *)
Stm_A_Rev_Axis000_Power(Enable := NOT M9999, Axis := Stm_A_Rev_Axis000);
(* Rung 1: #A(左側)ステッピング反転モータ1 原点復帰・動作設定パラメータ *)
//MC_HomeWithParameterの原点復帰パラメータ設定
//添付画像の参考値を設定（タッチパネルとの連携は未実装）
//実機使用前に原点信号・方向・速度・軸の単位を確認する
//このSTだけでは原点復帰を開始しない
//このST実行時は以下の固定値で上書きする

//原点復帰方式：近傍退避・原点近傍入力ON
Homing_Para_Stm.HomingMode := _mcHomeSwTurnHomeSwOn;
//原点入力：Z相（実機の信号対応を要確認）
Homing_Para_Stm.HomeInput := _mcZPhase;
//原点復帰の開始方向：負方向
Homing_Para_Stm.StartDir := _mcNegativeDirection;
//原点入力の検出方向：負方向
Homing_Para_Stm.HomeDir := _mcNegativeDirection;
//正側リミット入力時：即停止して反転
Homing_Para_Stm.PosiLmtMode := _mcRevImmediateStop;
//負側リミット入力時：即停止して反転
Homing_Para_Stm.NegaLmtMode := _mcRevImmediateStop;

//原点復帰速度 [指令単位/s]
Homing_Para_Stm.Vel := LREAL#40;
//原点近傍での接近速度 [指令単位/s]
Homing_Para_Stm.ApproachVel := LREAL#1;
//原点復帰の加速度 [指令単位/s^2]
Homing_Para_Stm.Acc := LREAL#100;
//原点復帰の減速度 [指令単位/s^2]
Homing_Para_Stm.Dec := LREAL#200;
//ジャーク [指令単位/s^3]：0はジャーク制御なし
Homing_Para_Stm.Jerk := LREAL#0;

//原点入力マスク距離 [指令単位]：今回の方式では未使用
Homing_Para_Stm.Mask := LREAL#0;
//原点確定後の現在位置 [指令単位]
Homing_Para_Stm.Offset := LREAL#0;
//押当て時間 [ms]：今回の方式では未使用
Homing_Para_Stm.PushTime := UINT#0;
//原点検出後の補正移動量 [指令単位]：0は補正移動なし
Homing_Para_Stm.Compensation := LREAL#0;
//原点補正移動時の速度 [指令単位/s]
Homing_Para_Stm.CompensationVel := LREAL#10;
(* Rung 2: 原点復帰完了 *)
Stm_A_Rev_Axis000_HomeWithParameter(Execute := Stm_A_Rev_Axis000_Origin AND Stm_A_Rev_Axis000_Power.Enable, Axis := Stm_A_Rev_Axis000, HomingParameter := Homing_Para_Stm);
Stm_A_Rev_Axis000_ZeroSet(Execute := Stm_A_Rev_Axis000_HomeWithParameter.Done, Axis := Stm_A_Rev_Axis000, Position := LREAL#0, ReferenceType := _eMC_REFERENCE_TYPE#_mcCommand);
Stm_A_Rev_Axis000_OriginDone := (Stm_A_Rev_Axis000_ZeroSet.Done OR Stm_A_Rev_Axis000_OriginDone) AND NOT M9999;

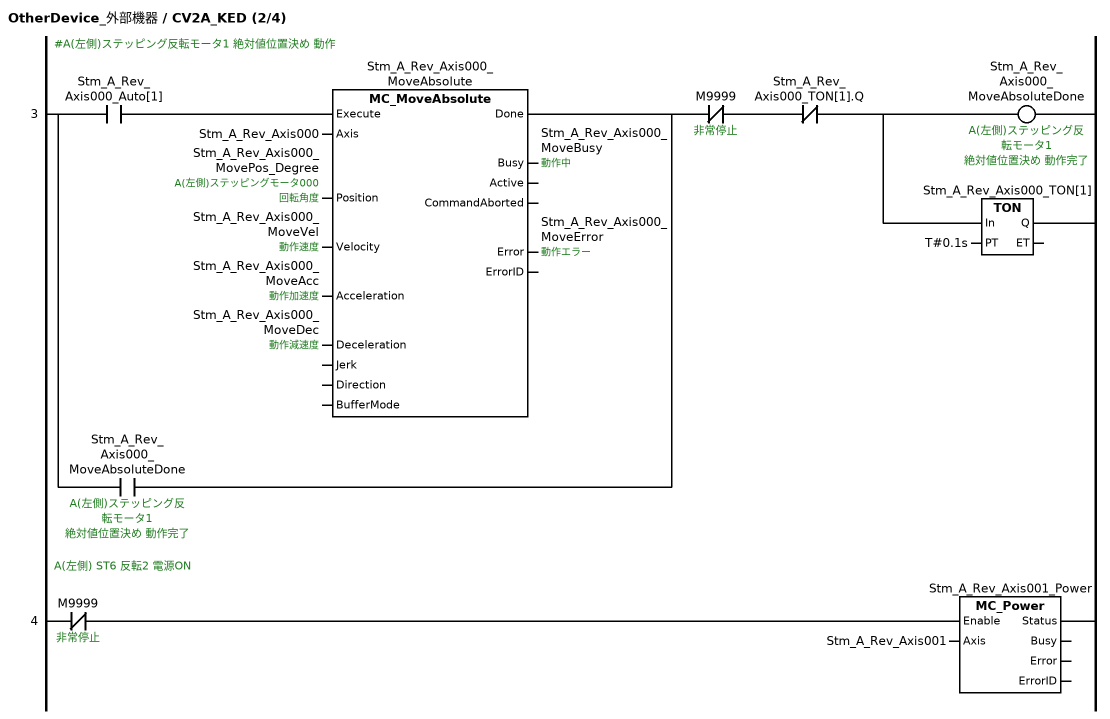
(* Rung 3: #A(左側)ステッピング反転モータ1 絶対値位置決め 動作 *)
Stm_A_Rev_Axis000_MoveAbsolute(Execute := Stm_A_Rev_Axis000_Auto[1], Axis := Stm_A_Rev_Axis000, Position := Stm_A_Rev_Axis000_MovePos_Degree, Velocity := Stm_A_Rev_Axis000_MoveVel, Acceleration := Stm_A_Rev_Axis000_MoveAcc, Deceleration := Stm_A_Rev_Axis000_MoveDec, Busy => Stm_A_Rev_Axis000_MoveBusy, Error => Stm_A_Rev_Axis000_MoveError);
_p51 := (Stm_A_Rev_Axis000_MoveAbsolute.Done OR Stm_A_Rev_Axis000_MoveAbsoluteDone) AND NOT M9999 AND NOT Stm_A_Rev_Axis000_TON[1].Q;
Stm_A_Rev_Axis000_MoveAbsoluteDone := _p51;
Stm_A_Rev_Axis000_TON[1](In := _p51, PT := T#0.1s);
(* Rung 4: A(左側) ST6 反転2 電源ON *)
Stm_A_Rev_Axis001_Power(Enable := NOT M9999, Axis := Stm_A_Rev_Axis001);

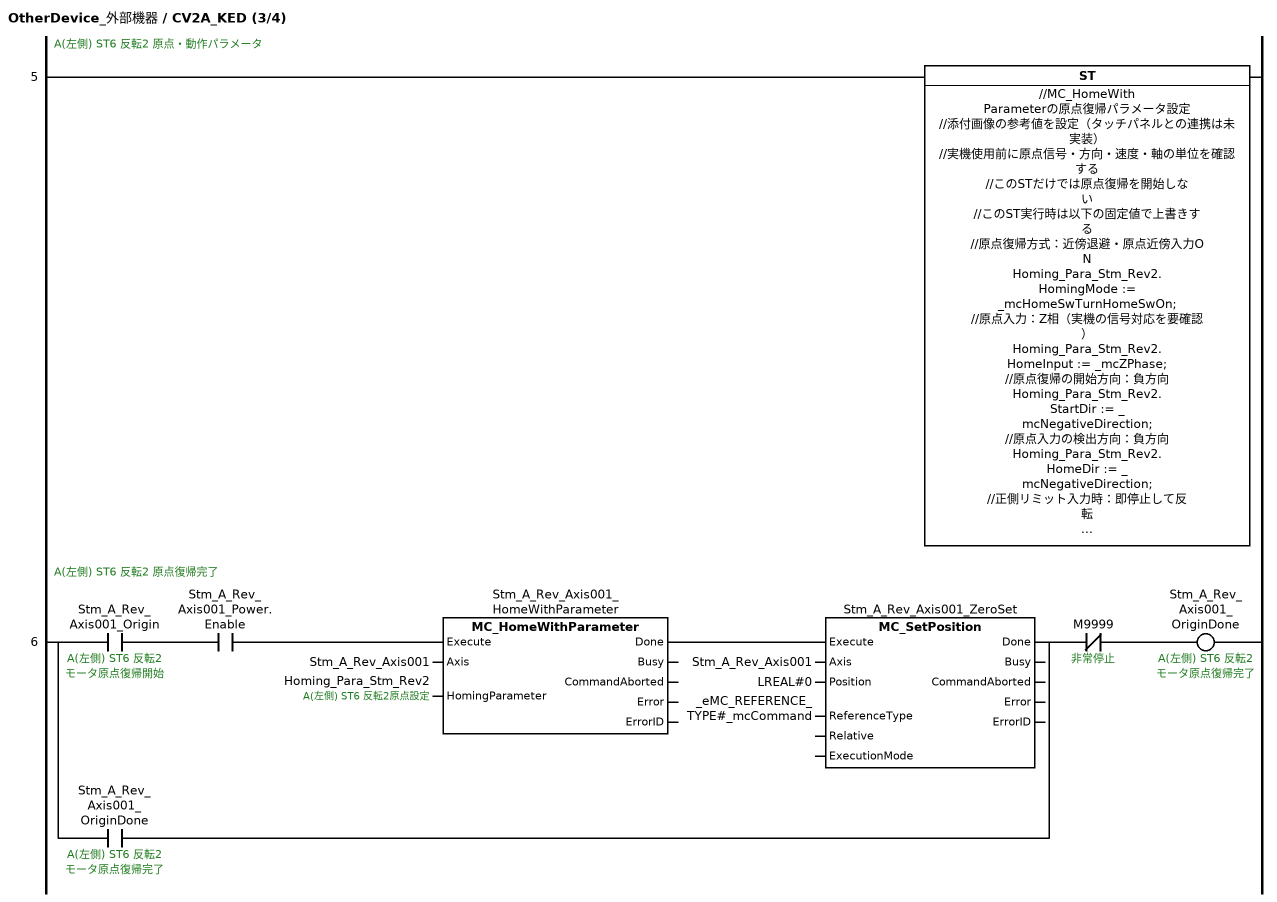
(* Rung 5: A(左側) ST6 反転2 原点・動作パラメータ *)
//MC_HomeWithParameterの原点復帰パラメータ設定
//添付画像の参考値を設定（タッチパネルとの連携は未実装）
//実機使用前に原点信号・方向・速度・軸の単位を確認する
//このSTだけでは原点復帰を開始しない
//このST実行時は以下の固定値で上書きする

//原点復帰方式：近傍退避・原点近傍入力ON
Homing_Para_Stm_Rev2.HomingMode := _mcHomeSwTurnHomeSwOn;
//原点入力：Z相（実機の信号対応を要確認）
Homing_Para_Stm_Rev2.HomeInput := _mcZPhase;
//原点復帰の開始方向：負方向
Homing_Para_Stm_Rev2.StartDir := _mcNegativeDirection;
//原点入力の検出方向：負方向
Homing_Para_Stm_Rev2.HomeDir := _mcNegativeDirection;
//正側リミット入力時：即停止して反転
Homing_Para_Stm_Rev2.PosiLmtMode := _mcRevImmediateStop;
//負側リミット入力時：即停止して反転
Homing_Para_Stm_Rev2.NegaLmtMode := _mcRevImmediateStop;

//原点復帰速度 [指令単位/s]
Homing_Para_Stm_Rev2.Vel := LREAL#40;
//原点近傍での接近速度 [指令単位/s]
Homing_Para_Stm_Rev2.ApproachVel := LREAL#1;
//原点復帰の加速度 [指令単位/s^2]
Homing_Para_Stm_Rev2.Acc := LREAL#100;
//原点復帰の減速度 [指令単位/s^2]
Homing_Para_Stm_Rev2.Dec := LREAL#200;
//ジャーク [指令単位/s^3]：0はジャーク制御なし
Homing_Para_Stm_Rev2.Jerk := LREAL#0;

//原点入力マスク距離 [指令単位]：今回の方式では未使用
Homing_Para_Stm_Rev2.Mask := LREAL#0;
//原点確定後の現在位置 [指令単位]
Homing_Para_Stm_Rev2.Offset := LREAL#0;
//押当て時間 [ms]：今回の方式では未使用
Homing_Para_Stm_Rev2.PushTime := UINT#0;
//原点検出後の補正移動量 [指令単位]：0は補正移動なし
Homing_Para_Stm_Rev2.Compensation := LREAL#0;
//原点補正移動時の速度 [指令単位/s]
Homing_Para_Stm_Rev2.CompensationVel := LREAL#10;
(* Rung 6: A(左側) ST6 反転2 原点復帰完了 *)
Stm_A_Rev_Axis001_HomeWithParameter(Execute := Stm_A_Rev_Axis001_Origin AND Stm_A_Rev_Axis001_Power.Enable, Axis := Stm_A_Rev_Axis001, HomingParameter := Homing_Para_Stm_Rev2);
Stm_A_Rev_Axis001_ZeroSet(Execute := Stm_A_Rev_Axis001_HomeWithParameter.Done, Axis := Stm_A_Rev_Axis001, Position := LREAL#0, ReferenceType := _eMC_REFERENCE_TYPE#_mcCommand);
Stm_A_Rev_Axis001_OriginDone := (Stm_A_Rev_Axis001_ZeroSet.Done OR Stm_A_Rev_Axis001_OriginDone) AND NOT M9999;

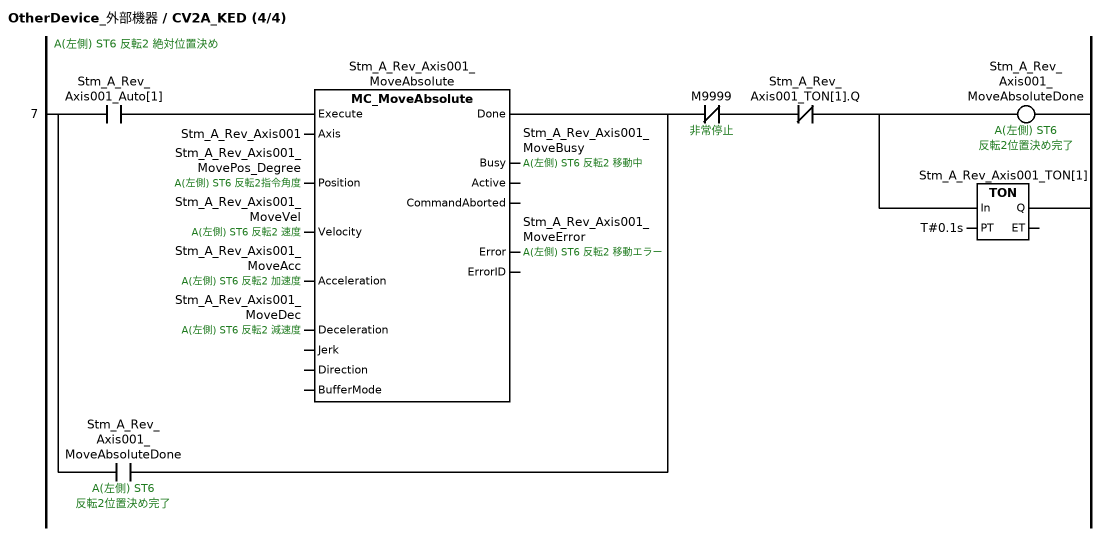
(* Rung 7: A(左側) ST6 反転2 絶対位置決め *)
Stm_A_Rev_Axis001_MoveAbsolute(Execute := Stm_A_Rev_Axis001_Auto[1], Axis := Stm_A_Rev_Axis001, Position := Stm_A_Rev_Axis001_MovePos_Degree, Velocity := Stm_A_Rev_Axis001_MoveVel, Acceleration := Stm_A_Rev_Axis001_MoveAcc, Deceleration := Stm_A_Rev_Axis001_MoveDec, Busy => Stm_A_Rev_Axis001_MoveBusy, Error => Stm_A_Rev_Axis001_MoveError);
_p52 := (Stm_A_Rev_Axis001_MoveAbsolute.Done OR Stm_A_Rev_Axis001_MoveAbsoluteDone) AND NOT M9999 AND NOT Stm_A_Rev_Axis001_TON[1].Q;
Stm_A_Rev_Axis001_MoveAbsoluteDone := _p52;
Stm_A_Rev_Axis001_TON[1](In := _p52, PT := T#0.1s);

(* Section HMI: ladder, written here as Structured Text *)

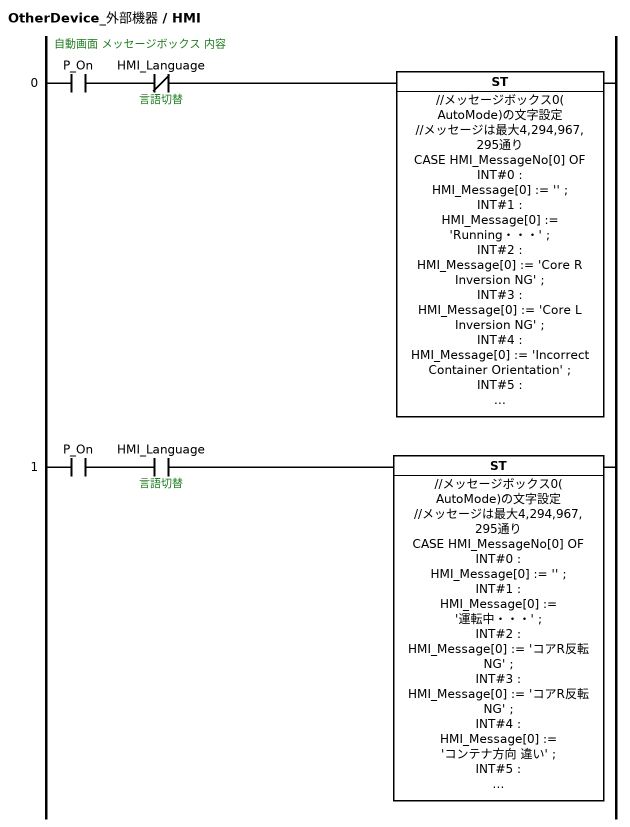
(* Rung 0: 自動画面 メッセージボックス 内容 *)
IF P_On AND NOT HMI_Language THEN
    //メッセージボックス0(AutoMode)の文字設定
    //メッセージは最大4,294,967,295通り
    	
    	CASE HMI_MessageNo[0] OF
    	
    	INT#0 :
    	HMI_Message[0] := '' ;
        INT#1 :
    	HMI_Message[0] := 'Running・・・' ;
    	INT#2 :
    	HMI_Message[0] := 'Core R Inversion NG' ;
    	INT#3 :
    	HMI_Message[0] := 'Core L Inversion NG' ;
    	INT#4 :
    	HMI_Message[0] := 'Incorrect Container Orientation' ;
    	INT#5 :
    	HMI_Message[0] := 'Packed Container Full' ;
         INT#6 :
    	HMI_Message[0] := 'No Container Added' ;
    	INT#7 :
    	HMI_Message[0] := 'Paused・・・' ;
        INT#8 :
    	HMI_Message[0] := 'R Stock Holder Qty Error' ;
    	INT#9 :
    	HMI_Message[0] := 'L Stock Holder Qty Error' ;
        INT#10 :
    	HMI_Message[0] := 'Step Running・・・' ;
    	INT#11 :
    	HMI_Message[0] := 'Work Discharge Complete' ;
    	INT#12 :
    	HMI_Message[0] := 'SD Error' ;
    	END_CASE;		
    	
END_IF;
(* Rung 1 *)
IF P_On AND HMI_Language THEN
    //メッセージボックス0(AutoMode)の文字設定
    //メッセージは最大4,294,967,295通り
    	
    	CASE HMI_MessageNo[0] OF
    	
    	INT#0 :
    	HMI_Message[0] := '' ;
    	INT#1 :
    	HMI_Message[0] := '運転中・・・' ;	
    	INT#2 :
    	HMI_Message[0] := 'コアR反転 NG' ;	
        INT#3 :
    	HMI_Message[0] := 'コアR反転 NG' ;
    	INT#4 :
    	HMI_Message[0] := 'コンテナ方向 違い' ;
    	INT#5 :
    	HMI_Message[0] := '梱包済みコンテナ 満杯 or 排出詰まり' ;
        INT#6 :
    	HMI_Message[0] := 'コンテナ 無 追加してください' ;
        INT#7 :
    	HMI_Message[0] := '一時停止中・・・' ;
        INT#8 :
    	HMI_Message[0] := '右ストックフォルダ 入数ミス 取り除いて 再スタート' ;
        INT#9 :
    	HMI_Message[0] := '左ストックフォルダ 入数ミス 取り除いて 再スタート' ;
    	INT#10 :
    	HMI_Message[0] := 'ステップ運転中・・・' ;
    	INT#11 :
    	HMI_Message[0] := 'ワーク排出完了' ;
    	INT#12 :
    	HMI_Message[0] := 'SDカードエラー' ;
    	END_CASE;		
    	
END_IF;
END_PROGRAM

